(* IEC 61131-3 sources: NachHouse_TST/API/api_V12, 8 files *)

(* ---- _01_Types.ST ---- *)
// Konštanty určujú rozmery virtuálnej pamäte a počet typov ; Constants define virtual-memory dimensions and the number of data types.
VAR_GLOBAL CONSTANT
  _NH_ZONES {HIDDEN} : USINT := 5;      // Počet podporovaných pamäťových zón PLC ; Number of PLC memory zones used by this model.
  _NH_RAM {HIDDEN}   : UDINT := 10000;  // Veľkosť poľa mRam v bajtoch ; Size of the mRam byte array.
  _NH_CFG {HIDDEN}   : INT := 2;        // Počet typov registrovaných v aCfg ; Number of data types registered in aCfg.
END_VAR

// Nasledujú interné typy, dátové záznamy a dve publikované aplikačné štruktúry ; The following are internal types, data records, and two published application structures.
TYPE
  // Príznaky štartu a inicializácie programu ; Program startup and initialization flags.
  NH_SYS {HIDDEN}: STRUCT
    Ini     : INT := 250;    // Hodnota 250 povoľuje jednorazové naplnenie testovacích dát ; Value 250 enables the one-time test-data initialization.
    Restart : BOOL := TRUE;  // Označuje, že PLC práve štartuje ; Indicates that the PLC is starting.
  END_STRUCT;
  // Príklad spoločných identifikačných polí v oboch typoch ; Example of shared identification fields in both data types.
  NH_CFG_ALL {HIDDEN}: STRUCT
    RoomID     : INT := 12;  // Ukážkové ID miestnosti v spoločnej časti ; Sample room ID in the shared section.
    CategoryID : INT := 23;  // Ukážkové ID kategórie v spoločnej časti ; Sample category ID in the shared section.
  END_STRUCT;
  // Metaúdaje jedného typu: kód, veľkosť, počet viet a umiestnenie v mRam ; Metadata for one type: code, size, record count, and location in mRam.
  NH_CFG: STRUCT
    cfg     : STRING[4];                    // Kód typu, veľkosť vety, adresa, offset v mRam a počet viet ; Type code, record size, address, mRam offset, and record count.
    Siz     : UDINT;
    Ram     : UDINT;
    iRam    : UDINT;
    Rec     : UDINT;
    par     : USINT;                        // Pomocné klasifikačné a referenčné metadáta typu ; Auxiliary type classification and reference metadata.
    cat     : USINT;
    ref     : USINT := 251;
    ver     : USINT;
    tGrp    : USINT;                        // Klasifikačné údaje a veľkosti konfiguračnej/spoločnej časti ; Classification values and configuration/shared-section sizes.
    al      : USINT;
    cx      : UDINT;
    cf      : USINT := SIZEOF(NH_CFG_ALL);
    me      : UDINT;                        // Veľkosť stavovej časti, HW/I/O údaje a príznaky použiteľnosti ; State-section size, hardware/I/O data, and validity flags.
    hw      : USINT;
    io      : UDINT;
    Enabled : BOOL;
    ok      : BOOL;
  END_STRUCT;
  // Spoločné polia hlavičky každého záznamu ; Shared header fields for every record.
  NH_REC_ALL {HIDDEN}: STRUCT
    Ok : BOOL := TRUE;  // Príznak platnosti záznamu ; Record-validity flag.
    ID : INT;           // Identifikátor záznamu ; Record identifier.
  END_STRUCT;
  // Premenné živého stavu miestnosti uložené v časti mem ; Live room-state fields stored in the mem section.
  NH_ROOM_MEM: STRUCT
    rec          : NH_REC_ALL;  // Hlavička vety a spoločné identifikačné údaje ; Record header and shared identification data.
    all          : NH_CFG_ALL;
    Temperature  : REAL;        // Testovacie merania a stavové príznaky miestnosti ; Test measurements and room-state flags.
    Humidity     : REAL;
    Presence     : BOOL;
    DayPhase     : UINT;
    CategoryMask : DWORD;       // Maska kategórií, alarm a ďalšie binárne príznaky stavu ; Category mask, alarm level, and additional Boolean state flags.
    AlarmLevel   : USINT;
    Online       : BOOL;
    Twilight     : BOOL;
  END_STRUCT;
  // Konfiguračná časť miestnosti ; testovacie polia pokrývajú rôzne IEC typy ; Room configuration ; test fields cover different IEC data types.
  NH_ROOM_CFG: STRUCT
    Name           : STRING[32];                              // Názov a testovacie celé čísla so znamienkom aj bez neho ; Name and signed/unsigned integer test values.
    _Dint          : DINT;
    _Sint          : SINT;
    _Usint         : USINT;
    _Uint          : UINT;                                    // Testovacie 16-bitové a plávajúce čísla a krátky reťazec ; 16-bit and floating-point test values plus a short string.
    _Real          : REAL;
    _LReal         : LREAL;
    _String        : STRING[30];
    _StringCZSK    : STRING := 'SVKBEGIN_+ľščťžýáíé_SVKEND';  // Reťazec s diakritikou overuje prevod CP1250 na UTF-8 a späť ; A diacritic-bearing string tests conversion between CP1250 and UTF-8.
    _BYTE          : BYTE;                                    // Testovacie bajtové a časové typy ; Byte-sized and date/time test types.
    _WORD          : WORD;
    _TIME          : TIME;
    _DATE          : DATE;
    _TIME_OF_DAY   : TOD;                                     // Testovacie typy času dňa a dátumu s časom ; Test values for time-of-day and date-time types.
    _DATE_AND_TIME : DT;
  END_STRUCT;
  // Celá verejná veta miestnosti spája živý stav a konfiguráciu ; One public room record combines live state and configuration.
  NH_ROOM {PUBLIC}: STRUCT
    mem : NH_ROOM_MEM;  // Podštruktúra prevádzkového stavu miestnosti ; Nested room operating-state structure.
    cfg : NH_ROOM_CFG;  // Podštruktúra konfiguračných hodnôt miestnosti ; Nested room-configuration structure.
  END_STRUCT;
  // Živý stav používateľa oddelený od jeho konfigurácie ; Live user state separated from user configuration.
  NH_USERS_MEM: STRUCT
    rec        : NH_REC_ALL;  // Hlavička, spoločné identifikátory a stav pripojenia ; Header, shared identifiers, and connection state.
    all        : NH_CFG_ALL;
    Connected  : BOOL;
    LastError  : STRING[80];  // Posledná chyba a časová značka poslednej aktualizácie ; Last error and timestamp of the latest update.
    LastUpdate : UDINT;
  END_STRUCT;
  // Konfigurácia používateľa vrátane práv, zón, IP a ďalších polí ; User configuration including rights, zones, IP addresses, and other fields.
  NH_USERS_CFG: STRUCT
    Name       : STRING[32];                                                                                                              // Meno používateľa a predvoľby úvodnej obrazovky ; User name and home-screen preferences.
    LoginHome  : BOOL := TRUE;
    DshSet     : BOOL := FALSE;
    OwnDSH     : BOOL := TRUE;                                                                                                            // Príznaky vlastných obrazoviek a úroveň oprávnenia ; Custom-screen flags and access-right level.
    OwnQCK     : BOOL := TRUE;
    UsrRight   : USINT := 1;
    ZonList    : ARRAY[1..16] OF BOOL := [1, 1, 1, 1, 1, 1, 1, 1, 1, 1, 1, 1, 1, 1, 1, 1];                                                // Prístup používateľa k šestnástim zónam ; User access flags for sixteen zones.
    sbj        : USINT := 1;                                                                                                              // Predmet, jazyk a osem obľúbených položiek ; Subject, language, and eight favorites.
    lng        : USINT;
    fav        : ARRAY[0..7] OF USINT;
    keyPas     : STRING[6];                                                                                                               // Krátky testovací kľúč, počet IP adries a tri adresy ; Test key, IP-address count, and three addresses.
    IPnbr      : USINT := 1;
    IP         : ARRAY[1..3] OF STRING[15];
    mail       : STRING[50];                                                                                                              // Kontaktný e-mail a testovacie autorizačné tokeny ; Contact email and test authorization tokens.
    TOKENAPPLE : STRING[90];
    TOKENUNI   : STRING[100];
    gsm        : STRING[15];                                                                                                              // Telefón, vzhľad a osem príznakov správ ; Phone, appearance, and eight message flags.
    skin       : USINT;
    msg        : ARRAY[0..7] OF BOOL;
    Brw        : ARRAY[0..30] OF USINT := [0, 1, 1, 1, 1, 1, 1, 1, 1, 1, 1, 1, 1, 1, 1, 1, 1, 1, 1, 1, 1, 1, 1, 1, 1, 1, 1, 1, 1, 1, 1];  // Tridsaťjeden testovacích hodnôt pre prehliadač ; Thirty-one test values for browser-related settings.
  END_STRUCT;
  // Celá verejná veta používateľa spája stav a konfiguráciu ; One public user record combines state and configuration.
  NH_USER {PUBLIC}: STRUCT
    mem : NH_USERS_MEM;
    cfg : NH_USERS_CFG;
  END_STRUCT;
END_TYPE

VAR_GLOBAL
  mRam : ARRAY[0.._NH_RAM] OF BYTE;        // Spoločný bajtový priestor, v ktorom sú uložené všetky vety ; Shared byte-addressable memory containing all records.
  aSys : NH_SYS;                           // Stavové príznaky inicializácie programu ; Program initialization state.
  aCfg : ARRAY[1.._NH_CFG] OF NH_CFG := [  // Tabuľka typov: určuje ich veľkosti, počty viet a rozloženie v mRam ; Type table: defines sizes, record counts, and placement in mRam.
    (cfg := 'ROOM', Enabled := TRUE, ver := 1, Siz := SIZEOF(NH_ROOM),
     Rec := 10, cx := SIZEOF(NH_ROOM.cfg), me := SIZEOF(NH_ROOM.mem)),
    (cfg := 'USER', Enabled := TRUE, ver := 1, Siz := SIZEOF(NH_USER),
     Rec := 10, cx := SIZEOF(NH_USER.cfg), me := SIZEOF(NH_USER.mem),
     cat := 31, ref := 254)
  ];
  xRoom : PTR_TO NH_ROOM;  // Ukazovateľ na začiatok poľa viet ROOM v mRam ; Pointer to the first ROOM record in mRam.
  xUser : PTR_TO NH_USER;  // Ukazovateľ na začiatok poľa viet USER v mRam ; Pointer to the first USER record in mRam.

  yRooms : ARRAY[1..10] OF NH_ROOM;  // Iba zdroj testovacích dát ; po skopírovaní do mRam sa ďalej nepoužíva. ; Test-data source only ; unused after copying into mRam.
  yUsers : ARRAY[1..10] OF NH_USER;  // Zdroj testovacích viet USER ; po skopírovaní do mRam sa ďalej nepoužíva ; Source of USER test records ; unused after copying into mRam.

  DepRq {PUBLIC_API}   : BOOL := FALSE;        // Požiadavka na aktiváciu balíka ; Package-activation request.
  DepRes {PUBLIC_API}  : USINT := 0;           // Výsledkový kód aktivácie balíka ; Package-activation result code.
  BuildNo {PUBLIC_API} : UDINT := 2026100726;  // Číslo zostavenia na kontrolu nasadenej verzie ; Build number used to verify the deployed version.

  TxCf {PUBLIC_API}   : USINT := 2;  // Klient nastaví typ a vetu ; TxRq ako posledné spustí export. Nula znamená všetky vety. ; The client sets type and record ; TxRq starts the export last. Zero means all records.
  TxRec {PUBLIC_API}  : UDINT := 0;  // Číslo exportovanej vety ; nula znamená všetky vety vybraného typu ; Record to export ; zero means all records of the selected type.
  TxRq {PUBLIC_API}   : UDINT := 1;  // Klient zmenou čísla spustí nový export ; A new value starts an export request.
  TxDone {PUBLIC_API} : UDINT := 0;  // Potvrdí číslo dokončenej požiadavky na export ; Echoes the completed export request number.
  TxErr {PUBLIC_API}  : USINT := 0;  // Nula znamená úspech ; nenulová hodnota označuje chybu exportu ; Zero means success ; nonzero indicates an export error.

  RxRq    {PUBLIC_API} : UDINT := 0;  // Po prijatí rx.json klient zapíše nové RxRq a tým spustí jeho import. ; After rx.json is received, the client writes a new RxRq to start its import.
  RxDone  {PUBLIC_API} : UDINT := 0;  // Potvrdí číslo dokončenej požiadavky na import ; Echoes the completed import request number.
  RxErr   {PUBLIC_API} : USINT := 0;  // Nula znamená úspešný import ; inak obsahuje kód chyby ; Zero means import succeeded ; otherwise contains an error code.

  rxBuf   {PUBLIC_API} : ARRAY[0..63] OF DWORD;  // Jeden blok klienta má 64 DWORD, teda kapacitu 256 bajtov. ; One client block contains 64 DWORD values, providing 256 bytes of capacity. ; Klient zapíše dáta a metadáta ; RbRq mení až po nich. ; The client writes data and metadata first, then changes RbRq.
  RbOfs   {PUBLIC_API} : UDINT := 0;             // Offset bloku v celom súbore ; Block offset within the complete file.
  RbLen   {PUBLIC_API} : UINT := 0;              // Počet platných bajtov v tomto bloku ; Number of valid bytes in this block.
  RbTotal {PUBLIC_API} : UDINT := 0;             // Celková veľkosť prijímaného súboru ; Total size of the incoming file.
  RbCrc   {PUBLIC_API} : DWORD := 0;             // Očakávaný CRC32 súčet celého súboru ; Expected CRC32 checksum of the complete file.
  RbRq    {PUBLIC_API} : UDINT := 0;             // Spúšťací čítač bloku ; klient ho zapisuje až po dátach ; Block trigger counter ; written only after the block data.
  RbAck   {PUBLIC_API} : UDINT := 0;             // Potvrdzuje spracované číslo bloku ; Acknowledges the processed block number.
  RbWrote {PUBLIC_API} : UDINT := 0;             // Počet bajtov už uložených do rx.json ; Number of bytes already written to rx.json.
  RbReady {PUBLIC_API} : BOOL := FALSE;          // TRUE znamená celý súbor uložený a CRC overené ; TRUE means the full file is written and its CRC is valid.
  RbErr   {PUBLIC_API} : USINT := 0;             // Výsledok posledného bloku ; nula znamená úspech ; Result of the latest block ; zero means success.
END_VAR

(* ---- _03_Schema.ST ---- *)
// Automaticky vygenerované z api_V12.pux ; neupravovať ručne. ; GENERATED from api_V12.pux. Do not edit manually.
VAR_GLOBAL CONSTANT
  SCH_BOOL          : USINT := 16#01;        // Kód typu BOOL v schéme ; BOOL type code in the schema
  SCH_SINT          : USINT := 16#02;        // Kód typu SINT v schéme ; SINT type code in the schema
  SCH_USINT         : USINT := 16#03;        // Kód typu USINT v schéme ; USINT type code in the schema
  SCH_INT           : USINT := 16#04;        // Kód typu INT v schéme ; INT type code in the schema
  SCH_UINT          : USINT := 16#05;        // Kód typu UINT v schéme ; UINT type code in the schema
  SCH_DINT          : USINT := 16#06;        // Kód typu DINT v schéme ; DINT type code in the schema
  SCH_UDINT         : USINT := 16#07;        // Kód typu UDINT v schéme ; UDINT type code in the schema
  SCH_BYTE          : USINT := 16#08;        // Kód typu BYTE v schéme ; BYTE type code in the schema
  SCH_WORD          : USINT := 16#09;        // Kód typu WORD v schéme ; WORD type code in the schema
  SCH_DWORD         : USINT := 16#0A;        // Kód typu DWORD v schéme ; DWORD type code in the schema
  SCH_REAL          : USINT := 16#0B;        // Kód typu REAL v schéme ; REAL type code in the schema
  SCH_LREAL         : USINT := 16#0C;        // Kód typu LREAL v schéme ; LREAL type code in the schema
  SCH_STRING        : USINT := 16#0D;        // Kód reťazca v schéme ; String type code in the schema
  SCH_TIME          : USINT := 16#0E;        // Kód typu TIME v schéme ; TIME type code in the schema
  SCH_DATE          : USINT := 16#0F;        // Kód typu DATE v schéme ; DATE type code in the schema
  SCH_TIME_OF_DAY   : USINT := 16#10;        // Kód typu TOD v schéme ; TOD type code in the schema
  SCH_DATE_AND_TIME : USINT := 16#11;        // Kód typu DT v schéme ; DT type code in the schema
  SCH_STRUCT        : USINT := 16#12;        // Kód vnorenej štruktúry v schéme ; Nested-structure type code in the schema
  SCH_ARRAY         : USINT := 16#80;        // Príznak poľa kombinovaný so základným typom ; Array flag combined with the base type
  SCH_BASE          : USINT := 16#7F;        // Maska na získanie základného typu ; Mask used to extract the base type
  SCH_DEF_N         : UINT := 2;             // Počet definovaných aplikačných typov ; Number of application types defined
  SCH_NODE_N        : UINT := 62;            // Počet uzlov stromu štruktúr ; Number of structure-tree nodes
  SCH_LEAF_N        : UINT := 115;           // Počet úplných ciest k položkám ; Number of complete field paths
  SCH_PUX_CRC       : DWORD := 16#B72908B3;  // Kontrolný súčet zdrojového PUX ; Checksum of the source PUX
END_VAR

TYPE
  NH_SCH : STRUCT
    Cfg  : USINT;       // Poradové číslo typu v aCfg ; Type index in aCfg
    Code : STRING[4];   // Kód typu používaný v JSON obálke ; Type code used in the JSON envelope
    Nam  : STRING[16];  // Názov typu alebo uzla podľa kontextu ; Type or node name, depending on context
    Siz  : UDINT;       // Veľkosť jednej celej vety v bajtoch ; Size of one complete record in bytes
    Fst  : UINT;        // Index prvého uzla typu ; Index of the first node for this type
    Cnt  : UINT;        // Počet uzlov typu ; Number of nodes for this type
    LFst : UINT;        // Index prvej úplnej cesty poľa ; Index of the first complete field path
    LCnt : UINT;        // Počet úplných ciest poľa ; Number of complete field paths
  END_STRUCT;
  NH_NODE : STRUCT
    Nam  : STRING[14];  // Názov typu alebo uzla podľa kontextu ; Type or node name, depending on context
    Tag  : USINT;       // Kód dátového typu a prípadný príznak poľa ; Data-type code and optional array flag
    Ofs  : UINT;        // Offset položky od začiatku rodiča ; Field offset from the parent start
    Span : UINT;        // Veľkosť položky v bajtoch ; Field size in bytes
    Aux  : UINT;        // Doplnkový údaj podľa typu uzla ; Auxiliary value interpreted by node type
    Cnt  : UINT;        // Počet uzlov typu ; Number of nodes for this type
    Lo   : INT;         // Dolná hranica poľa ; Array lower bound
  END_STRUCT;
  NH_LEAF : STRUCT
    Pth    : STRING[18];  // Úplná cesta poľa od koreňa vety ; Complete field path from the record root
    Tag    : USINT;       // Kód dátového typu a prípadný príznak poľa ; Data-type code and optional array flag
    Ofs    : UINT;        // Offset položky od začiatku rodiča ; Field offset from the parent start
    Span   : UINT;        // Veľkosť položky v bajtoch ; Field size in bytes
    BitPos : SINT;        // Pozícia BOOL poľa v bajte ; BOOL field bit position within its byte
  END_STRUCT;
END_TYPE

VAR_GLOBAL
  aSch : ARRAY[1..2] OF NH_SCH := [  // Tabuľka rozsahov uzlov a polí pre každý typ ; Per-type ranges of nodes and fields
    (Cfg := 1, Code := 'ROOM', Nam := 'NH_ROOM', Siz := 216, Fst := 1, Cnt := 31, LFst := 1, LCnt := 27),
    (Cfg := 2, Code := 'USER', Nam := 'NH_USER', Siz := 488, Fst := 32, Cnt := 31, LFst := 28, LCnt := 88)
  ];
  aNode : ARRAY[1..62] OF NH_NODE := [  // Sploštený strom všetkých uzlov štruktúr ; Flattened tree of all structure nodes
    (Nam := 'mem', Tag := 16#12, Ofs := 0, Span := 24, Aux := 14, Cnt := 0, Lo := 0),
    (Nam := 'rec', Tag := 16#12, Ofs := 0, Span := 3, Aux := 2, Cnt := 0, Lo := 0),
    (Nam := 'Ok', Tag := 16#01, Ofs := 0, Span := 1, Aux := 0, Cnt := 0, Lo := 0),
    (Nam := 'ID', Tag := 16#04, Ofs := 1, Span := 2, Aux := 0, Cnt := 0, Lo := 0),
    (Nam := 'all', Tag := 16#12, Ofs := 3, Span := 4, Aux := 2, Cnt := 0, Lo := 0),
    (Nam := 'RoomID', Tag := 16#04, Ofs := 0, Span := 2, Aux := 0, Cnt := 0, Lo := 0),
    (Nam := 'CategoryID', Tag := 16#04, Ofs := 2, Span := 2, Aux := 0, Cnt := 0, Lo := 0),
    (Nam := 'Temperature', Tag := 16#0B, Ofs := 7, Span := 4, Aux := 0, Cnt := 0, Lo := 0),
    (Nam := 'Humidity', Tag := 16#0B, Ofs := 11, Span := 4, Aux := 0, Cnt := 0, Lo := 0),
    (Nam := 'Presence', Tag := 16#01, Ofs := 15, Span := 1, Aux := 0, Cnt := 0, Lo := 0),
    (Nam := 'DayPhase', Tag := 16#05, Ofs := 16, Span := 2, Aux := 0, Cnt := 0, Lo := 0),
    (Nam := 'CategoryMask', Tag := 16#0A, Ofs := 18, Span := 4, Aux := 0, Cnt := 0, Lo := 0),
    (Nam := 'AlarmLevel', Tag := 16#03, Ofs := 22, Span := 1, Aux := 0, Cnt := 0, Lo := 0),
    (Nam := 'Online', Tag := 16#01, Ofs := 23, Span := 1, Aux := 0, Cnt := 0, Lo := 0),
    (Nam := 'Twilight', Tag := 16#01, Ofs := 23, Span := 1, Aux := 1, Cnt := 0, Lo := 0),
    (Nam := 'cfg', Tag := 16#12, Ofs := 24, Span := 192, Aux := 15, Cnt := 0, Lo := 0),
    (Nam := 'Name', Tag := 16#0D, Ofs := 0, Span := 33, Aux := 0, Cnt := 0, Lo := 0),
    (Nam := '_Dint', Tag := 16#06, Ofs := 33, Span := 4, Aux := 0, Cnt := 0, Lo := 0),
    (Nam := '_Sint', Tag := 16#02, Ofs := 37, Span := 1, Aux := 0, Cnt := 0, Lo := 0),
    (Nam := '_Usint', Tag := 16#03, Ofs := 38, Span := 1, Aux := 0, Cnt := 0, Lo := 0),
    (Nam := '_Uint', Tag := 16#05, Ofs := 39, Span := 2, Aux := 0, Cnt := 0, Lo := 0),
    (Nam := '_Real', Tag := 16#0B, Ofs := 41, Span := 4, Aux := 0, Cnt := 0, Lo := 0),
    (Nam := '_LReal', Tag := 16#0C, Ofs := 45, Span := 8, Aux := 0, Cnt := 0, Lo := 0),
    (Nam := '_String', Tag := 16#0D, Ofs := 53, Span := 31, Aux := 0, Cnt := 0, Lo := 0),
    (Nam := '_StringCZSK', Tag := 16#0D, Ofs := 84, Span := 81, Aux := 0, Cnt := 0, Lo := 0),
    (Nam := '_BYTE', Tag := 16#08, Ofs := 165, Span := 1, Aux := 0, Cnt := 0, Lo := 0),
    (Nam := '_WORD', Tag := 16#09, Ofs := 166, Span := 2, Aux := 0, Cnt := 0, Lo := 0),
    (Nam := '_TIME', Tag := 16#0E, Ofs := 168, Span := 4, Aux := 0, Cnt := 0, Lo := 0),
    (Nam := '_DATE', Tag := 16#0F, Ofs := 172, Span := 8, Aux := 0, Cnt := 0, Lo := 0),
    (Nam := '_TIME_OF_DAY', Tag := 16#10, Ofs := 180, Span := 4, Aux := 0, Cnt := 0, Lo := 0),
    (Nam := '_DATE_AND_TIME', Tag := 16#11, Ofs := 184, Span := 8, Aux := 0, Cnt := 0, Lo := 0),
    (Nam := 'mem', Tag := 16#12, Ofs := 0, Span := 93, Aux := 9, Cnt := 0, Lo := 0),
    (Nam := 'rec', Tag := 16#12, Ofs := 0, Span := 3, Aux := 2, Cnt := 0, Lo := 0),
    (Nam := 'Ok', Tag := 16#01, Ofs := 0, Span := 1, Aux := 0, Cnt := 0, Lo := 0),
    (Nam := 'ID', Tag := 16#04, Ofs := 1, Span := 2, Aux := 0, Cnt := 0, Lo := 0),
    (Nam := 'all', Tag := 16#12, Ofs := 3, Span := 4, Aux := 2, Cnt := 0, Lo := 0),
    (Nam := 'RoomID', Tag := 16#04, Ofs := 0, Span := 2, Aux := 0, Cnt := 0, Lo := 0),
    (Nam := 'CategoryID', Tag := 16#04, Ofs := 2, Span := 2, Aux := 0, Cnt := 0, Lo := 0),
    (Nam := 'Connected', Tag := 16#01, Ofs := 7, Span := 1, Aux := 0, Cnt := 0, Lo := 0),
    (Nam := 'LastError', Tag := 16#0D, Ofs := 8, Span := 81, Aux := 0, Cnt := 0, Lo := 0),
    (Nam := 'LastUpdate', Tag := 16#07, Ofs := 89, Span := 4, Aux := 0, Cnt := 0, Lo := 0),
    (Nam := 'cfg', Tag := 16#12, Ofs := 93, Span := 395, Aux := 20, Cnt := 0, Lo := 0),
    (Nam := 'Name', Tag := 16#0D, Ofs := 0, Span := 33, Aux := 0, Cnt := 0, Lo := 0),
    (Nam := 'LoginHome', Tag := 16#01, Ofs := 33, Span := 1, Aux := 0, Cnt := 0, Lo := 0),
    (Nam := 'DshSet', Tag := 16#01, Ofs := 33, Span := 1, Aux := 1, Cnt := 0, Lo := 0),
    (Nam := 'OwnDSH', Tag := 16#01, Ofs := 33, Span := 1, Aux := 2, Cnt := 0, Lo := 0),
    (Nam := 'OwnQCK', Tag := 16#01, Ofs := 33, Span := 1, Aux := 3, Cnt := 0, Lo := 0),
    (Nam := 'UsrRight', Tag := 16#03, Ofs := 34, Span := 1, Aux := 0, Cnt := 0, Lo := 0),
    (Nam := 'ZonList', Tag := 16#81, Ofs := 35, Span := 2, Aux := 0, Cnt := 16, Lo := 1),
    (Nam := 'sbj', Tag := 16#03, Ofs := 37, Span := 1, Aux := 0, Cnt := 0, Lo := 0),
    (Nam := 'lng', Tag := 16#03, Ofs := 38, Span := 1, Aux := 0, Cnt := 0, Lo := 0),
    (Nam := 'fav', Tag := 16#83, Ofs := 39, Span := 8, Aux := 1, Cnt := 8, Lo := 0),
    (Nam := 'keyPas', Tag := 16#0D, Ofs := 47, Span := 7, Aux := 0, Cnt := 0, Lo := 0),
    (Nam := 'IPnbr', Tag := 16#03, Ofs := 54, Span := 1, Aux := 0, Cnt := 0, Lo := 0),
    (Nam := 'IP', Tag := 16#8D, Ofs := 55, Span := 48, Aux := 16, Cnt := 3, Lo := 1),
    (Nam := 'mail', Tag := 16#0D, Ofs := 103, Span := 51, Aux := 0, Cnt := 0, Lo := 0),
    (Nam := 'TOKENAPPLE', Tag := 16#0D, Ofs := 154, Span := 91, Aux := 0, Cnt := 0, Lo := 0),
    (Nam := 'TOKENUNI', Tag := 16#0D, Ofs := 245, Span := 101, Aux := 0, Cnt := 0, Lo := 0),
    (Nam := 'gsm', Tag := 16#0D, Ofs := 346, Span := 16, Aux := 0, Cnt := 0, Lo := 0),
    (Nam := 'skin', Tag := 16#03, Ofs := 362, Span := 1, Aux := 0, Cnt := 0, Lo := 0),
    (Nam := 'msg', Tag := 16#81, Ofs := 363, Span := 1, Aux := 0, Cnt := 8, Lo := 0),
    (Nam := 'Brw', Tag := 16#83, Ofs := 364, Span := 31, Aux := 1, Cnt := 31, Lo := 0)
  ];
  aLeaf : ARRAY[1..115] OF NH_LEAF := [  // Tabuľka úplných názvov koncových polí ; Lookup table of complete leaf-field names
    (Pth := 'mem.rec.Ok', Tag := 16#01, Ofs := 0, Span := 1, BitPos := 0),
    (Pth := 'mem.rec.ID', Tag := 16#04, Ofs := 1, Span := 2, BitPos := -1),
    (Pth := 'mem.all.RoomID', Tag := 16#04, Ofs := 3, Span := 2, BitPos := -1),
    (Pth := 'mem.all.CategoryID', Tag := 16#04, Ofs := 5, Span := 2, BitPos := -1),
    (Pth := 'mem.Temperature', Tag := 16#0B, Ofs := 7, Span := 4, BitPos := -1),
    (Pth := 'mem.Humidity', Tag := 16#0B, Ofs := 11, Span := 4, BitPos := -1),
    (Pth := 'mem.Presence', Tag := 16#01, Ofs := 15, Span := 1, BitPos := 0),
    (Pth := 'mem.DayPhase', Tag := 16#05, Ofs := 16, Span := 2, BitPos := -1),
    (Pth := 'mem.CategoryMask', Tag := 16#0A, Ofs := 18, Span := 4, BitPos := -1),
    (Pth := 'mem.AlarmLevel', Tag := 16#03, Ofs := 22, Span := 1, BitPos := -1),
    (Pth := 'mem.Online', Tag := 16#01, Ofs := 23, Span := 1, BitPos := 0),
    (Pth := 'mem.Twilight', Tag := 16#01, Ofs := 23, Span := 1, BitPos := 1),
    (Pth := 'cfg.Name', Tag := 16#0D, Ofs := 24, Span := 33, BitPos := -1),
    (Pth := 'cfg._Dint', Tag := 16#06, Ofs := 57, Span := 4, BitPos := -1),
    (Pth := 'cfg._Sint', Tag := 16#02, Ofs := 61, Span := 1, BitPos := -1),
    (Pth := 'cfg._Usint', Tag := 16#03, Ofs := 62, Span := 1, BitPos := -1),
    (Pth := 'cfg._Uint', Tag := 16#05, Ofs := 63, Span := 2, BitPos := -1),
    (Pth := 'cfg._Real', Tag := 16#0B, Ofs := 65, Span := 4, BitPos := -1),
    (Pth := 'cfg._LReal', Tag := 16#0C, Ofs := 69, Span := 8, BitPos := -1),
    (Pth := 'cfg._String', Tag := 16#0D, Ofs := 77, Span := 31, BitPos := -1),
    (Pth := 'cfg._StringCZSK', Tag := 16#0D, Ofs := 108, Span := 81, BitPos := -1),
    (Pth := 'cfg._BYTE', Tag := 16#08, Ofs := 189, Span := 1, BitPos := -1),
    (Pth := 'cfg._WORD', Tag := 16#09, Ofs := 190, Span := 2, BitPos := -1),
    (Pth := 'cfg._TIME', Tag := 16#0E, Ofs := 192, Span := 4, BitPos := -1),
    (Pth := 'cfg._DATE', Tag := 16#0F, Ofs := 196, Span := 8, BitPos := -1),
    (Pth := 'cfg._TIME_OF_DAY', Tag := 16#10, Ofs := 204, Span := 4, BitPos := -1),
    (Pth := 'cfg._DATE_AND_TIME', Tag := 16#11, Ofs := 208, Span := 8, BitPos := -1),
    (Pth := 'mem.rec.Ok', Tag := 16#01, Ofs := 0, Span := 1, BitPos := 0),
    (Pth := 'mem.rec.ID', Tag := 16#04, Ofs := 1, Span := 2, BitPos := -1),
    (Pth := 'mem.all.RoomID', Tag := 16#04, Ofs := 3, Span := 2, BitPos := -1),
    (Pth := 'mem.all.CategoryID', Tag := 16#04, Ofs := 5, Span := 2, BitPos := -1),
    (Pth := 'mem.Connected', Tag := 16#01, Ofs := 7, Span := 1, BitPos := 0),
    (Pth := 'mem.LastError', Tag := 16#0D, Ofs := 8, Span := 81, BitPos := -1),
    (Pth := 'mem.LastUpdate', Tag := 16#07, Ofs := 89, Span := 4, BitPos := -1),
    (Pth := 'cfg.Name', Tag := 16#0D, Ofs := 93, Span := 33, BitPos := -1),
    (Pth := 'cfg.LoginHome', Tag := 16#01, Ofs := 126, Span := 1, BitPos := 0),
    (Pth := 'cfg.DshSet', Tag := 16#01, Ofs := 126, Span := 1, BitPos := 1),
    (Pth := 'cfg.OwnDSH', Tag := 16#01, Ofs := 126, Span := 1, BitPos := 2),
    (Pth := 'cfg.OwnQCK', Tag := 16#01, Ofs := 126, Span := 1, BitPos := 3),
    (Pth := 'cfg.UsrRight', Tag := 16#03, Ofs := 127, Span := 1, BitPos := -1),
    (Pth := 'cfg.ZonList[0]', Tag := 16#01, Ofs := 128, Span := 1, BitPos := 0),
    (Pth := 'cfg.ZonList[1]', Tag := 16#01, Ofs := 128, Span := 1, BitPos := 1),
    (Pth := 'cfg.ZonList[2]', Tag := 16#01, Ofs := 128, Span := 1, BitPos := 2),
    (Pth := 'cfg.ZonList[3]', Tag := 16#01, Ofs := 128, Span := 1, BitPos := 3),
    (Pth := 'cfg.ZonList[4]', Tag := 16#01, Ofs := 128, Span := 1, BitPos := 4),
    (Pth := 'cfg.ZonList[5]', Tag := 16#01, Ofs := 128, Span := 1, BitPos := 5),
    (Pth := 'cfg.ZonList[6]', Tag := 16#01, Ofs := 128, Span := 1, BitPos := 6),
    (Pth := 'cfg.ZonList[7]', Tag := 16#01, Ofs := 128, Span := 1, BitPos := 7),
    (Pth := 'cfg.ZonList[8]', Tag := 16#01, Ofs := 129, Span := 1, BitPos := 0),
    (Pth := 'cfg.ZonList[9]', Tag := 16#01, Ofs := 129, Span := 1, BitPos := 1),
    (Pth := 'cfg.ZonList[10]', Tag := 16#01, Ofs := 129, Span := 1, BitPos := 2),
    (Pth := 'cfg.ZonList[11]', Tag := 16#01, Ofs := 129, Span := 1, BitPos := 3),
    (Pth := 'cfg.ZonList[12]', Tag := 16#01, Ofs := 129, Span := 1, BitPos := 4),
    (Pth := 'cfg.ZonList[13]', Tag := 16#01, Ofs := 129, Span := 1, BitPos := 5),
    (Pth := 'cfg.ZonList[14]', Tag := 16#01, Ofs := 129, Span := 1, BitPos := 6),
    (Pth := 'cfg.ZonList[15]', Tag := 16#01, Ofs := 129, Span := 1, BitPos := 7),
    (Pth := 'cfg.sbj', Tag := 16#03, Ofs := 130, Span := 1, BitPos := -1),
    (Pth := 'cfg.lng', Tag := 16#03, Ofs := 131, Span := 1, BitPos := -1),
    (Pth := 'cfg.fav[0]', Tag := 16#03, Ofs := 132, Span := 1, BitPos := -1),
    (Pth := 'cfg.fav[1]', Tag := 16#03, Ofs := 133, Span := 1, BitPos := -1),
    (Pth := 'cfg.fav[2]', Tag := 16#03, Ofs := 134, Span := 1, BitPos := -1),
    (Pth := 'cfg.fav[3]', Tag := 16#03, Ofs := 135, Span := 1, BitPos := -1),
    (Pth := 'cfg.fav[4]', Tag := 16#03, Ofs := 136, Span := 1, BitPos := -1),
    (Pth := 'cfg.fav[5]', Tag := 16#03, Ofs := 137, Span := 1, BitPos := -1),
    (Pth := 'cfg.fav[6]', Tag := 16#03, Ofs := 138, Span := 1, BitPos := -1),
    (Pth := 'cfg.fav[7]', Tag := 16#03, Ofs := 139, Span := 1, BitPos := -1),
    (Pth := 'cfg.keyPas', Tag := 16#0D, Ofs := 140, Span := 7, BitPos := -1),
    (Pth := 'cfg.IPnbr', Tag := 16#03, Ofs := 147, Span := 1, BitPos := -1),
    (Pth := 'cfg.IP[0]', Tag := 16#0D, Ofs := 148, Span := 16, BitPos := -1),
    (Pth := 'cfg.IP[1]', Tag := 16#0D, Ofs := 164, Span := 16, BitPos := -1),
    (Pth := 'cfg.IP[2]', Tag := 16#0D, Ofs := 180, Span := 16, BitPos := -1),
    (Pth := 'cfg.mail', Tag := 16#0D, Ofs := 196, Span := 51, BitPos := -1),
    (Pth := 'cfg.TOKENAPPLE', Tag := 16#0D, Ofs := 247, Span := 91, BitPos := -1),
    (Pth := 'cfg.TOKENUNI', Tag := 16#0D, Ofs := 338, Span := 101, BitPos := -1),
    (Pth := 'cfg.gsm', Tag := 16#0D, Ofs := 439, Span := 16, BitPos := -1),
    (Pth := 'cfg.skin', Tag := 16#03, Ofs := 455, Span := 1, BitPos := -1),
    (Pth := 'cfg.msg[0]', Tag := 16#01, Ofs := 456, Span := 1, BitPos := 0),
    (Pth := 'cfg.msg[1]', Tag := 16#01, Ofs := 456, Span := 1, BitPos := 1),
    (Pth := 'cfg.msg[2]', Tag := 16#01, Ofs := 456, Span := 1, BitPos := 2),
    (Pth := 'cfg.msg[3]', Tag := 16#01, Ofs := 456, Span := 1, BitPos := 3),
    (Pth := 'cfg.msg[4]', Tag := 16#01, Ofs := 456, Span := 1, BitPos := 4),
    (Pth := 'cfg.msg[5]', Tag := 16#01, Ofs := 456, Span := 1, BitPos := 5),
    (Pth := 'cfg.msg[6]', Tag := 16#01, Ofs := 456, Span := 1, BitPos := 6),
    (Pth := 'cfg.msg[7]', Tag := 16#01, Ofs := 456, Span := 1, BitPos := 7),
    (Pth := 'cfg.Brw[0]', Tag := 16#03, Ofs := 457, Span := 1, BitPos := -1),
    (Pth := 'cfg.Brw[1]', Tag := 16#03, Ofs := 458, Span := 1, BitPos := -1),
    (Pth := 'cfg.Brw[2]', Tag := 16#03, Ofs := 459, Span := 1, BitPos := -1),
    (Pth := 'cfg.Brw[3]', Tag := 16#03, Ofs := 460, Span := 1, BitPos := -1),
    (Pth := 'cfg.Brw[4]', Tag := 16#03, Ofs := 461, Span := 1, BitPos := -1),
    (Pth := 'cfg.Brw[5]', Tag := 16#03, Ofs := 462, Span := 1, BitPos := -1),
    (Pth := 'cfg.Brw[6]', Tag := 16#03, Ofs := 463, Span := 1, BitPos := -1),
    (Pth := 'cfg.Brw[7]', Tag := 16#03, Ofs := 464, Span := 1, BitPos := -1),
    (Pth := 'cfg.Brw[8]', Tag := 16#03, Ofs := 465, Span := 1, BitPos := -1),
    (Pth := 'cfg.Brw[9]', Tag := 16#03, Ofs := 466, Span := 1, BitPos := -1),
    (Pth := 'cfg.Brw[10]', Tag := 16#03, Ofs := 467, Span := 1, BitPos := -1),
    (Pth := 'cfg.Brw[11]', Tag := 16#03, Ofs := 468, Span := 1, BitPos := -1),
    (Pth := 'cfg.Brw[12]', Tag := 16#03, Ofs := 469, Span := 1, BitPos := -1),
    (Pth := 'cfg.Brw[13]', Tag := 16#03, Ofs := 470, Span := 1, BitPos := -1),
    (Pth := 'cfg.Brw[14]', Tag := 16#03, Ofs := 471, Span := 1, BitPos := -1),
    (Pth := 'cfg.Brw[15]', Tag := 16#03, Ofs := 472, Span := 1, BitPos := -1),
    (Pth := 'cfg.Brw[16]', Tag := 16#03, Ofs := 473, Span := 1, BitPos := -1),
    (Pth := 'cfg.Brw[17]', Tag := 16#03, Ofs := 474, Span := 1, BitPos := -1),
    (Pth := 'cfg.Brw[18]', Tag := 16#03, Ofs := 475, Span := 1, BitPos := -1),
    (Pth := 'cfg.Brw[19]', Tag := 16#03, Ofs := 476, Span := 1, BitPos := -1),
    (Pth := 'cfg.Brw[20]', Tag := 16#03, Ofs := 477, Span := 1, BitPos := -1),
    (Pth := 'cfg.Brw[21]', Tag := 16#03, Ofs := 478, Span := 1, BitPos := -1),
    (Pth := 'cfg.Brw[22]', Tag := 16#03, Ofs := 479, Span := 1, BitPos := -1),
    (Pth := 'cfg.Brw[23]', Tag := 16#03, Ofs := 480, Span := 1, BitPos := -1),
    (Pth := 'cfg.Brw[24]', Tag := 16#03, Ofs := 481, Span := 1, BitPos := -1),
    (Pth := 'cfg.Brw[25]', Tag := 16#03, Ofs := 482, Span := 1, BitPos := -1),
    (Pth := 'cfg.Brw[26]', Tag := 16#03, Ofs := 483, Span := 1, BitPos := -1),
    (Pth := 'cfg.Brw[27]', Tag := 16#03, Ofs := 484, Span := 1, BitPos := -1),
    (Pth := 'cfg.Brw[28]', Tag := 16#03, Ofs := 485, Span := 1, BitPos := -1),
    (Pth := 'cfg.Brw[29]', Tag := 16#03, Ofs := 486, Span := 1, BitPos := -1),
    (Pth := 'cfg.Brw[30]', Tag := 16#03, Ofs := 487, Span := 1, BitPos := -1)
  ];
END_VAR

(* ---- _04_SchemaRun.ST ---- *)
// Stav validácie generovanej schémy ; Validation state for the generated schema.
VAR_GLOBAL
  SchOk    : BOOL := FALSE;  // TRUE až po úspešnej kontrole celej tabuľky schémy ; TRUE only after the entire schema table passes validation.
  SchErr   : USINT := 0;     // Kód prvej chyby zistený pri kontrole schémy ; First error code detected during schema validation.
  SchState : USINT := 0;     // Kontrola schémy sa vykoná raz a jej výsledok sa zapamätá ; Schema validation runs once and its result is cached. 0=new, 1=valid, 2=error
END_VAR

// Porovná vygenerovanú schému s aCfg a aktuálnym rozložením mRam. ; Compare the generated schema with aCfg and the current mRam layout.
// Overí počty, veľkosti, uzly a rozsahy schémy ešte pred prevodom ; Validate schema counts, sizes, nodes, and bounds before conversion.
FUNCTION SchInit : BOOL
  VAR
    Cf       : INT;                   // Index dátového typu v aCfg/aSch ; Data-type index in aCfg/aSch.
    Nd       : UINT;                  // Index práve kontrolovaného uzla štruktúry ; Index of the structure node being checked.
    Last     : UINT;                  // Posledný uzol patriaci aktuálnemu typu ; Last node belonging to the current type.
    Expected : UINT := 1;             // Očakávaný začiatok ďalšieho súvislého rozsahu uzlov ; Expected start of the next contiguous node range.
    BaseTag  : USINT;                 // Základný typ uzla po odobratí príznaku ARRAY ; Node base type after removing the ARRAY flag. ; Základný typ určuje výpočet prvku poľa ; The base type determines array-element addressing.
    NodeEnd  : UINT;                  // Koniec podstromu vnoreného STRUCT ; End of a nested STRUCT subtree.
    ElemSpan : UINT;                  // Veľkosť jedného prvku poľa STRUCT ; Size of one STRUCT-array element.
    Depth    : USINT;                 // Aktuálna hĺbka vnorenia pri kontrole uzlov ; Current nesting depth while validating nodes.
    EndStk   : ARRAY[0..15] OF UINT;  // Zásobník hraníc uzlov vnorených štruktúr ; Stack of node-range ends for nested structures.
    SpanStk  : ARRAY[0..15] OF UINT;  // Zásobník veľkostí rodičovských pamäťových oblastí ; Stack of parent memory-span sizes.
    RamEnd   : UDINT;                 // Koniec vyhradenej oblasti typu v mRam ; End of this type's reserved region in mRam.
  END_VAR

  SchInit := FALSE;
  // Použije zapamätaný úspech bez opakovania úplnej kontroly ; Reuse the cached success without repeating full validation.
  IF SchState = 1 THEN SchInit := TRUE; RETURN; END_IF;
  // Po predchádzajúcej chybe sa prevod bezpečne zastaví ; Stop conversion after a previously detected schema error.
  IF SchState = 2 THEN RETURN; END_IF;

  SchOk := FALSE;
  SchErr := 1;
  SchState := 2;
  IF SCH_DEF_N <> INT_TO_UINT(_NH_CFG) THEN RETURN; END_IF;

  // Porovná každý typ schémy s jeho konfiguráciou a rozložením v pamäti ; Compare each schema type with its configuration and memory layout.
  FOR Cf := 1 TO _NH_CFG DO
    IF aSch[Cf].Cfg <> INT_TO_USINT(Cf) THEN SchErr := 2; RETURN; END_IF;
    IF aSch[Cf].Code <> aCfg[Cf].cfg THEN SchErr := 3; RETURN; END_IF;
    IF aSch[Cf].Siz <> aCfg[Cf].Siz THEN SchErr := 4; RETURN; END_IF;
    IF (aSch[Cf].Fst <> Expected) OR (aSch[Cf].Cnt = 0) THEN SchErr := 5; RETURN; END_IF;
    Last := aSch[Cf].Fst + aSch[Cf].Cnt - 1;
    IF Last > SCH_NODE_N THEN SchErr := 6; RETURN; END_IF;
    Expected := Last + 1;

    RamEnd := aCfg[Cf].iRam + aCfg[Cf].Siz * aCfg[Cf].Rec;
    IF RamEnd > SIZEOF(mRam) THEN SchErr := 7; RETURN; END_IF;
    IF aCfg[Cf].Ram <> PTR_TO_UDINT(ADR(mRam[aCfg[Cf].iRam])) THEN SchErr := 8; RETURN; END_IF;

    Depth := 0;  // Začne kontrolu stromu uzlov od koreňa aktuálneho typu ; Start validating the node tree at the current type's root.
    EndStk[0] := Last + 1;
    SpanStk[0] := UDINT_TO_UINT(aSch[Cf].Siz);
    FOR Nd := aSch[Cf].Fst TO Last DO
      WHILE (Depth > 0) AND (Nd >= EndStk[Depth]) DO Depth := Depth - 1; END_WHILE;
      IF UINT_TO_UDINT(aNode[Nd].Ofs) + UINT_TO_UDINT(aNode[Nd].Span) > UINT_TO_UDINT(SpanStk[Depth]) THEN
        SchErr := 9; RETURN;
      END_IF;

      BaseTag := aNode[Nd].Tag MOD SCH_ARRAY;  // Oddelí základný dátový typ od príznaku poľa ; Separate the base data type from the array flag.
      IF (BaseTag < SCH_BOOL) OR (BaseTag > SCH_STRUCT) OR (aNode[Nd].Span = 0) THEN
        SchErr := 10; RETURN;
      END_IF;

      IF aNode[Nd].Tag >= SCH_ARRAY THEN
        IF aNode[Nd].Cnt = 0 THEN SchErr := 11; RETURN; END_IF;
        IF BaseTag = SCH_STRUCT THEN
          IF (aNode[Nd].Span MOD aNode[Nd].Cnt) <> 0 THEN SchErr := 12; RETURN; END_IF;
        ELSIF BaseTag = SCH_BOOL THEN
          IF (aNode[Nd].Aux + aNode[Nd].Cnt + 7) / 8 > aNode[Nd].Span THEN SchErr := 13; RETURN; END_IF;
        ELSE
          IF (aNode[Nd].Aux = 0) OR (aNode[Nd].Aux * aNode[Nd].Cnt <> aNode[Nd].Span) THEN
            SchErr := 14; RETURN;
          END_IF;
        END_IF;
      ELSE
        IF aNode[Nd].Cnt <> 0 THEN SchErr := 15; RETURN; END_IF;
        IF (BaseTag = SCH_BOOL) AND (aNode[Nd].Aux > 7) THEN SchErr := 16; RETURN; END_IF;
      END_IF;

      IF BaseTag = SCH_STRUCT THEN
        NodeEnd := Nd + 1 + aNode[Nd].Aux;
        IF NodeEnd > EndStk[Depth] THEN SchErr := 17; RETURN; END_IF;
        IF aNode[Nd].Aux > 0 THEN
          IF Depth >= 15 THEN SchErr := 18; RETURN; END_IF;
          IF aNode[Nd].Tag >= SCH_ARRAY THEN ElemSpan := aNode[Nd].Span / aNode[Nd].Cnt;
          ELSE ElemSpan := aNode[Nd].Span;
          END_IF;
          Depth := Depth + 1;
          EndStk[Depth] := NodeEnd;
          SpanStk[Depth] := ElemSpan;
        END_IF;
      END_IF;
    END_FOR;
  END_FOR;

  IF Expected <> SCH_NODE_N + 1 THEN SchErr := 19; RETURN; END_IF;
  SchErr := 0;  // Všetky kontroly prešli ; SchInit môže povoliť prevod ; All checks passed ; SchInit may allow conversion.
  SchOk := TRUE;
  SchState := 1;
  SchInit := TRUE;
END_FUNCTION

// Vráti začiatok zvolenej vety v mRam ; Rec sa čísluje od 1. ; Return the selected record's base address in mRam ; Rec is one-based.
// Vráti adresu vybranej vety v mRam alebo nulu pri neplatnom výbere ; Return the selected record's mRam address, or zero for an invalid selection.
FUNCTION SchRoot : UDINT
  VAR_INPUT
    Cf  : USINT;
    Rec : UDINT;
  END_VAR
  SchRoot := 0;
  IF NOT SchInit() THEN RETURN; END_IF;
  IF (Cf < 1) OR (Cf > UINT_TO_USINT(SCH_DEF_N)) THEN RETURN; END_IF;
  IF (Rec < 1) OR (Rec > aCfg[Cf].Rec) THEN RETURN; END_IF;
  IF NOT aCfg[Cf].Enabled OR NOT aCfg[Cf].ok THEN RETURN; END_IF;
  SchRoot := aCfg[Cf].Ram + (Rec - 1) * aCfg[Cf].Siz;
END_FUNCTION

// Vypočíta adresu uzla v rodičovi ; El pri poli je skutočný IEC index. ; Calculate a node address within its parent ; El is the actual IEC array index.
// Vypočíta adresu položky alebo prvku poľa z rodičovskej adresy a offsetu ; Calculate a field/array-element address from its parent and offset.
FUNCTION SchAdr : UDINT
  VAR_INPUT
    Parent : UDINT;
    Nd     : UINT;   // Index práve kontrolovaného uzla štruktúry ; Index of the structure node being checked.
    El     : INT;
  END_VAR
  VAR
    BaseTag : USINT;  // Základný typ uzla po odobratí príznaku ARRAY ; Node base type after removing the ARRAY flag. ; Základný typ určuje výpočet prvku poľa ; The base type determines array-element addressing.
    K       : UINT;   // Poradové číslo prvku od dolnej hranice poľa ; Zero-based element index from the array lower bound.
    BitPos  : UINT;   // Bitová pozícia BOOL prvku v bajte ; Bit position of a BOOL element within its byte.
  END_VAR
  SchAdr := 0;
  IF NOT SchInit() OR (Parent = 0) OR (Nd < 1) OR (Nd > SCH_NODE_N) THEN RETURN; END_IF;
  IF aNode[Nd].Tag < SCH_ARRAY THEN
    SchAdr := Parent + UINT_TO_UDINT(aNode[Nd].Ofs);
    RETURN;
  END_IF;
  IF (El < aNode[Nd].Lo) OR (El >= aNode[Nd].Lo + UINT_TO_INT(aNode[Nd].Cnt)) THEN RETURN; END_IF;
  K := INT_TO_UINT(El - aNode[Nd].Lo);
  BaseTag := aNode[Nd].Tag MOD SCH_ARRAY;
  IF BaseTag = SCH_BOOL THEN
    BitPos := aNode[Nd].Aux + K;
    SchAdr := Parent + UINT_TO_UDINT(aNode[Nd].Ofs) + UINT_TO_UDINT(BitPos / 8);
  ELSIF BaseTag = SCH_STRUCT THEN
    SchAdr := Parent + UINT_TO_UDINT(aNode[Nd].Ofs) + UINT_TO_UDINT(K * (aNode[Nd].Span / aNode[Nd].Cnt));
  ELSE
    SchAdr := Parent + UINT_TO_UDINT(aNode[Nd].Ofs) + UINT_TO_UDINT(K * aNode[Nd].Aux);
  END_IF;
END_FUNCTION

// Vráti bitovú pozíciu BOOL ; pri ostatných typoch vráti -1. ; Return the BOOL bit position, or -1 for other types.
// Vráti bitovú pozíciu BOOL ; pri inom type vráti -1 ; Return a BOOL bit position, or -1 for another type.
FUNCTION SchBit : SINT
  VAR_INPUT
    Nd : UINT;  // Index práve kontrolovaného uzla štruktúry ; Index of the structure node being checked.
    El : INT;
  END_VAR
  VAR
    K : UINT;  // Poradové číslo prvku od dolnej hranice poľa ; Zero-based element index from the array lower bound.
  END_VAR
  SchBit := -1;
  IF (Nd < 1) OR (Nd > SCH_NODE_N) THEN RETURN; END_IF;
  IF (aNode[Nd].Tag MOD SCH_ARRAY) <> SCH_BOOL THEN RETURN; END_IF;
  IF aNode[Nd].Tag < SCH_ARRAY THEN
    SchBit := UINT_TO_SINT(aNode[Nd].Aux);
    RETURN;
  END_IF;
  IF (El < aNode[Nd].Lo) OR (El >= aNode[Nd].Lo + UINT_TO_INT(aNode[Nd].Cnt)) THEN RETURN; END_IF;
  K := INT_TO_UINT(El - aNode[Nd].Lo);
  SchBit := UINT_TO_SINT((aNode[Nd].Aux + K) MOD 8);
END_FUNCTION

// Nájde ďalší uzol rovnakej úrovne a preskočí vnorený STRUCT. ; Find the next node at the same level, skipping a nested STRUCT.
// Vráti nasledujúci súrodenecký uzol a preskočí vnorený podstrom ; Return the next sibling node, skipping any nested subtree.
FUNCTION SchNext : UINT
  VAR_INPUT
    Nd : UINT;
  END_VAR
  SchNext := 0;
  IF (Nd < 1) OR (Nd > SCH_NODE_N) THEN RETURN; END_IF;
  IF (aNode[Nd].Tag MOD SCH_ARRAY) = SCH_STRUCT THEN SchNext := Nd + 1 + aNode[Nd].Aux;
  ELSE SchNext := Nd + 1;
  END_IF;
END_FUNCTION

(* ---- _05_TxJson.ST ---- *)
VAR_GLOBAL
  TxPath    : STRING[80] := '//RAM/tx.json';     // Cieľový súbor exportovaného JSON ; Destination file for exported JSON
  TxLogPath : STRING[80] := '//RAM/tx.log';      // Súbor meraní exportu ; Export measurement log file
  TxCRLF    : STRING[2] := '$0D$0A';             // Koniec riadka používaný v súbore ; Line ending used in the file
  TxH       : HANDLE := INVALID_HANDLE_VALUE;    // Handle otvoreného exportného súboru ; Handle of the open export file
  TxSeen    : UDINT := 0;                        // Posledná požiadavka už spracovaná PLC ; Latest request already processed by the PLC
  TxWorkErr : USINT := 0;                        // Pracovný kód chyby exportu ; Working export error code
  TxBytes   : UDINT := 0;                        // Počet bajtov zapísaných do súboru ; Number of bytes written to the file
  TxHex     : STRING[16] := '0123456789ABCDEF';  // Tabuľka číslic na zápis hexadecimálnych hodnôt ; Digit table for hexadecimal output
  TxSt      : USINT := 0;                        // Stavový automat exportu ; Export state-machine state
  TxCfW     : USINT := 0;                        // Typ vybraný pre aktuálny export ; Type selected for the current export
  TxFrom    : UDINT := 0;                        // Prvé číslo exportovanej vety ; First record number to export
  TxTo      : UDINT := 0;                        // Posledné číslo exportovanej vety ; Last record number to export
  TxNow     : UDINT := 0;                        // Číslo vety spracúvanej teraz ; Record number currently being processed
  TxRqW     : UDINT := 0;                        // Číslo požiadavky aktuálneho exportu ; Request number for the current export
  TxMode    : USINT := 0;                        // Režim výberu viet ; Record-selection mode ; 1=one, 2=range, 3=all
  TxMs0     : UDINT := 0;                        // Čas začiatku exportu v milisekundách ; Export start time in milliseconds
  TxMs1     : UDINT := 0;                        // Čas konca exportu v milisekundách ; Export end time in milliseconds
  TxDur     : UDINT := 0;                        // Trvanie exportu v milisekundách ; Export duration in milliseconds
  TxCyc     : UDINT := 0;                        // Počítadlo cyklov PLC ; PLC-cycle counter
  TxCyc0    : UDINT := 0;                        // Počítadlo cyklov pri štarte exportu ; PLC-cycle count at export start
  TxCycN    : UDINT := 0;                        // Počet cyklov spotrebovaných exportom ; Number of cycles used by the export
  TxDoneN   : UDINT := 0;                        // Počet dokončených viet ; Number of completed records
END_VAR

// Zapíše ľubovoľný úsek pamäte do otvoreného JSON súboru a kontroluje počet bajtov. ; Write a raw memory span to the open JSON file and verify the byte count.
FUNCTION TxWriteRaw : BOOL
  VAR_INPUT
    Pos : UDINT;  // Začiatočná adresa alebo offset zapisovaných dát ; Start address or offset of the data being written
    Siz : UDINT;  // Počet bajtov zapisovaného úseku ; Number of bytes in the section being written
  END_VAR
  VAR
    N : UDINT;  // Počet bajtov skutočne zapísaných funkciou ; Number of bytes actually written by the function
  END_VAR
  TxWriteRaw := FALSE;
  IF Siz = 0 THEN TxWriteRaw := TRUE; RETURN; END_IF;
  N := FileWrite(hFile := TxH, adrBuf := Pos, size := Siz);
  TxBytes := TxBytes + N;
  IF N <> Siz THEN TxWorkErr := 3; RETURN; END_IF;
  TxWriteRaw := TRUE;
END_FUNCTION

// Zapíše textový reťazec do exportného súboru. ; Write a text string to the export file.
FUNCTION TxWrite : BOOL
  VAR_INPUT
    Text : STRING[255];  // Textový obsah zapisovaný do JSON ; Text content being written to JSON
  END_VAR
  TxWrite := TxWriteRaw(Pos := PTR_TO_UDINT(ADR(Text)), Siz := INT_TO_UDINT(LEN(Text)));
END_FUNCTION

// Zapíše text medzi úvodzovky JSON. ; Write text enclosed in JSON quotes.
FUNCTION TxWriteQuoted : BOOL
  VAR_INPUT
    Text : STRING[255];  // Textový obsah zapisovaný do JSON ; Text content being written to JSON
  END_VAR
  TxWriteQuoted := FALSE;
  IF NOT TxWrite(Text := '"') THEN RETURN; END_IF;
  IF NOT TxWrite(Text := Text) THEN RETURN; END_IF;
  IF NOT TxWrite(Text := '"') THEN RETURN; END_IF;
  TxWriteQuoted := TRUE;
END_FUNCTION

// Prevedie reťazec PLC z CP1250 na UTF-8 a escapuje riadiace znaky JSON. ; Convert the PLC string from CP1250 to UTF-8 and escape JSON control characters.
// Prevedie PLC reťazec na korektný UTF-8 reťazec JSON. ; Convert a PLC string into valid UTF-8 JSON text.
// Skopíruje pevný úsek PLC STRING, prevedie CP1250 na UTF-8 a začne JSON reťazec. ; Copy a fixed PLC STRING span, convert CP1250 to UTF-8, and open a JSON string.
FUNCTION TxWriteString : BOOL
  VAR_INPUT
    Pos  : UDINT;  // Začiatočná adresa alebo offset zapisovaných dát ; Start address or offset of the data being written
    Span : UINT;   // Veľkosť hodnoty podľa schémy ; Value size from the schema
  END_VAR
  VAR
    Cp  : STRING[255];  // Počet bajtov v PLC reťazci ; Number of bytes in the PLC string
    Utf : STRING[255];  // Reťazec po prevode do UTF-8 ; String after conversion to UTF-8
    Src : PTR_TO BYTE;  // Ukazovateľ na zdrojové bajty ; Pointer to the source bytes
    P   : PTR_TO BYTE;  // Pracovný ukazovateľ na hodnotu ; Working pointer to the value
    H   : PTR_TO BYTE;  // Hexadecimálna číslica ; Hexadecimal digit
    Q   : PTR_TO BYTE;  // Pracovný znak pri escapovaní JSON ; Working character during JSON escaping
    B   : BYTE;         // Pracovný bajt hodnoty ; Working value byte
    N   : UDINT;        // Počet bajtov skutočne zapísaných funkciou ; Number of bytes actually written by the function
    I   : UINT;         // Index opakovania alebo poľa ; Loop or array index
    J   : UINT;         // Druhý index vnoreného prechodu ; Secondary index for nested traversal
  END_VAR
  TxWriteString := FALSE;
  IF (Span = 0) OR (Span > SIZEOF(Cp)) THEN TxWorkErr := 7; RETURN; END_IF;
  Cp := '';
  Utf := '';
  Src := UDINT_TO_PTR(Pos);
  N := MemCpyPtr(source := Src, dest := ADR(Cp), length := UINT_TO_UDINT(Span));
  IF N <> UINT_TO_UDINT(Span) THEN TxWorkErr := 7; RETURN; END_IF;
  N := CP1250_TO_UTF8(cp1250 := Cp, utf8 := Utf, maxLen := 255);
  IF (Cp <> '') AND (N = 0) THEN TxWorkErr := 7; RETURN; END_IF;
  IF NOT TxWrite(Text := '"') THEN RETURN; END_IF;
  P := ADR(Utf);
  H := ADR(TxHex);
  // Každý UTF-8 bajt zapíše priamo alebo ho escapuje podľa pravidiel JSON. ; Write each UTF-8 byte directly or escape it according to JSON rules.
  FOR I := 1 TO INT_TO_UINT(LEN(Utf)) DO
    B := P^;
    CASE B OF
      8:  IF NOT TxWrite(Text := '\b') THEN RETURN; END_IF;
      9:  IF NOT TxWrite(Text := '\t') THEN RETURN; END_IF;
      10: IF NOT TxWrite(Text := '\n') THEN RETURN; END_IF;
      12: IF NOT TxWrite(Text := '\f') THEN RETURN; END_IF;
      13: IF NOT TxWrite(Text := '\r') THEN RETURN; END_IF;
      34: IF NOT TxWrite(Text := '\"') THEN RETURN; END_IF;
      92: IF NOT TxWrite(Text := '\\') THEN RETURN; END_IF;
      ELSE
        IF B < 32 THEN
          IF NOT TxWrite(Text := '\u00') THEN RETURN; END_IF;
          Q := H;
          J := 0;
          WHILE J < BYTE_TO_UINT(B) / 16 DO Q := Q + 1; J := J + 1; END_WHILE;
          IF NOT TxWriteRaw(Pos := PTR_TO_UDINT(Q), Siz := 1) THEN RETURN; END_IF;
          Q := H;
          J := 0;
          WHILE J < BYTE_TO_UINT(B) MOD 16 DO Q := Q + 1; J := J + 1; END_WHILE;
          IF NOT TxWriteRaw(Pos := PTR_TO_UDINT(Q), Siz := 1) THEN RETURN; END_IF;
        ELSE
          IF NOT TxWriteRaw(Pos := PTR_TO_UDINT(P), Siz := 1) THEN RETURN; END_IF;
        END_IF;
    END_CASE;
    P := P + 1;
  END_FOR;
  IF NOT TxWrite(Text := '"') THEN RETURN; END_IF;
  TxWriteString := TRUE;
END_FUNCTION

// Načíta jednu hodnotu podľa typu v schéme a zapíše ju do JSON. ; Read one value according to its schema type and write it to JSON.
// Schéma dodá typ a adresu ; nižšie sa hodnota prečíta cez ukazovateľ správneho typu. ; The schema supplies type and address ; the value is read through a correctly typed pointer.
FUNCTION TxWriteValue : BOOL
  VAR_INPUT
    Parent : UDINT;  // Adresa rodičovskej štruktúry v mRam ; Address of the parent structure in mRam
    Nd     : UINT;   // Index uzla aktuálnej položky schémy ; Schema-node index of the current field
    El     : INT;    // Index prvku poľa ; Array element index
  END_VAR
  VAR
    ValAdr : UDINT;         // Adresa hodnoty v mRam ; Address of the value in mRam
    Tag    : USINT;         // Základný typ hodnoty ; Base type of the value
    BitPos : SINT;          // Pozícia BOOL v bajte ; BOOL bit position within its byte
    Mask   : UINT;          // Maska na vyčítanie jedného BOOL bitu ; Mask used to read one BOOL bit
    I      : SINT;          // Index opakovania alebo poľa ; Loop or array index
    Text   : STRING[255];   // Textový obsah zapisovaný do JSON ; Text content being written to JSON
    PB     : PTR_TO BYTE;
    PS     : PTR_TO SINT;
    PU     : PTR_TO USINT;
    PI     : PTR_TO INT;
    PUI    : PTR_TO UINT;
    PDI    : PTR_TO DINT;
    PUD    : PTR_TO UDINT;
    PW     : PTR_TO WORD;
    PDW    : PTR_TO DWORD;
    PR     : PTR_TO REAL;
    PLR    : PTR_TO LREAL;
    PT     : PTR_TO TIME;
    PDate  : PTR_TO DATE;
    PTod   : PTR_TO TOD;
    PDT    : PTR_TO DT;
  END_VAR
  TxWriteValue := FALSE;
  ValAdr := SchAdr(Parent := Parent, Nd := Nd, El := El);
  IF ValAdr = 0 THEN TxWorkErr := 6; RETURN; END_IF;
  Tag := aNode[Nd].Tag MOD SCH_ARRAY;

  // Vyberie prevod podľa IEC dátového typu položky. ; Select conversion according to the field's IEC data type.
  CASE Tag OF
    SCH_BOOL:
      PB := UDINT_TO_PTR(ValAdr);
      BitPos := SchBit(Nd := Nd, El := El);
      IF BitPos < 0 THEN TxWorkErr := 6; RETURN; END_IF;
      Mask := 1;
      FOR I := 1 TO BitPos DO Mask := Mask * 2; END_FOR;
      IF (BYTE_TO_UINT(PB^) / Mask) MOD 2 = 1 THEN Text := 'true'; ELSE Text := 'false'; END_IF;
    SCH_SINT: PS := UDINT_TO_PTR(ValAdr); Text := SINT_TO_STRING(PS^);
    SCH_USINT: PU := UDINT_TO_PTR(ValAdr); Text := USINT_TO_STRING(PU^);
    SCH_INT: PI := UDINT_TO_PTR(ValAdr); Text := INT_TO_STRING(PI^);
    SCH_UINT: PUI := UDINT_TO_PTR(ValAdr); Text := UINT_TO_STRING(PUI^);
    SCH_DINT: PDI := UDINT_TO_PTR(ValAdr); Text := DINT_TO_STRING(PDI^);
    SCH_UDINT: PUD := UDINT_TO_PTR(ValAdr); Text := UDINT_TO_STRING(PUD^);
    SCH_BYTE: PB := UDINT_TO_PTR(ValAdr); Text := UDINT_TO_STRING(BYTE_TO_UDINT(PB^));
    SCH_WORD: PW := UDINT_TO_PTR(ValAdr); Text := UDINT_TO_STRING(WORD_TO_UDINT(PW^));
    SCH_DWORD: PDW := UDINT_TO_PTR(ValAdr); Text := UDINT_TO_STRING(DWORD_TO_UDINT(PDW^));
    SCH_REAL: PR := UDINT_TO_PTR(ValAdr); Text := REAL_TO_STRING(PR^);
    SCH_LREAL: PLR := UDINT_TO_PTR(ValAdr); Text := LREAL_TO_STRING(PLR^);
    SCH_STRING:
      TxWriteValue := TxWriteString(Pos := ValAdr, Span := aNode[Nd].Span);
      RETURN;
    SCH_TIME: PT := UDINT_TO_PTR(ValAdr); Text := TIME_TO_STRING(PT^);
    SCH_DATE: PDate := UDINT_TO_PTR(ValAdr); Text := DATE_TO_STRING(PDate^);
    SCH_TIME_OF_DAY: PTod := UDINT_TO_PTR(ValAdr); Text := TOD_TO_STRING(PTod^);
    SCH_DATE_AND_TIME: PDT := UDINT_TO_PTR(ValAdr); Text := DT_TO_STRING(PDT^);
    ELSE TxWorkErr := 6; RETURN;
  END_CASE;

  IF (Tag = SCH_TIME) OR (Tag = SCH_DATE) OR (Tag = SCH_TIME_OF_DAY) OR (Tag = SCH_DATE_AND_TIME) THEN
    TxWriteValue := TxWriteQuoted(Text := Text);
  ELSE
    TxWriteValue := TxWrite(Text := Text);
  END_IF;
END_FUNCTION

// Prečíta PLC systémové hodiny v milisekundách pre meranie exportu. ; Read the PLC millisecond clock for export timing.
FUNCTION TxClockMs : UDINT
  VAR_EXTERNAL
    AT %SL52 : DWORD;
  END_VAR
  TxClockMs := DWORD_TO_UDINT(%SL52);
END_FUNCTION

// Zapíše jeden riadok do meracieho logu exportu. ; Write one line to the export measurement log.
FUNCTION TxLogPut : BOOL
  VAR_INPUT
    Hnd  : HANDLE;
    Text : STRING[255];  // Textový obsah zapisovaný do JSON ; Text content being written to JSON
  END_VAR
  VAR
    N : UDINT;  // Počet bajtov skutočne zapísaných funkciou ; Number of bytes actually written by the function
  END_VAR
  N := FileWrite(hFile := Hnd, adrBuf := PTR_TO_UDINT(ADR(Text)), size := INT_TO_UDINT(LEN(Text)));
  TxLogPut := N = INT_TO_UDINT(LEN(Text));
END_FUNCTION

// Zapíše parametre, výsledok a namerané trvanie exportu do tx.log. ; Write export parameters, result, and timing to tx.log.
FUNCTION TxWriteLog : BOOL
  VAR
    Hnd    : HANDLE;
    Line   : STRING[255];
    Closed : BOOL;          // Príznak úspešného uzatvorenia súboru ; Flag indicating the file closed successfully
    Ok     : BOOL := TRUE;  // Príznak úspešného zápisu ; Flag indicating a successful write
  END_VAR
  TxWriteLog := FALSE;
  Hnd := FileOpen(fileName := TxLogPath, mode := F_WRITE);
  IF Hnd = INVALID_HANDLE_VALUE THEN RETURN; END_IF;

  Line := CONCAT('api_V12 TX export', TxCRLF); Ok := Ok AND TxLogPut(Hnd := Hnd, Text := Line);
  Line := CONCAT('file=RAM/tx.json', TxCRLF); Ok := Ok AND TxLogPut(Hnd := Hnd, Text := Line);
  Line := CONCAT('rq=', UDINT_TO_STRING(TxRqW), TxCRLF); Ok := Ok AND TxLogPut(Hnd := Hnd, Text := Line);
  Line := CONCAT('cf=', USINT_TO_STRING(TxCfW), TxCRLF); Ok := Ok AND TxLogPut(Hnd := Hnd, Text := Line);
  IF (TxCfW >= 1) AND (TxCfW <= UINT_TO_USINT(SCH_DEF_N)) THEN
    Line := CONCAT('type=', aSch[TxCfW].Code, TxCRLF); Ok := Ok AND TxLogPut(Hnd := Hnd, Text := Line);
  END_IF;
  IF TxMode = 3 THEN Line := CONCAT('mode=all', TxCRLF);
  ELSIF TxMode = 2 THEN Line := CONCAT('mode=range', TxCRLF);
  ELSE Line := CONCAT('mode=one', TxCRLF);
  END_IF;
  Ok := Ok AND TxLogPut(Hnd := Hnd, Text := Line);
  Line := CONCAT('from=', UDINT_TO_STRING(TxFrom), TxCRLF); Ok := Ok AND TxLogPut(Hnd := Hnd, Text := Line);
  Line := CONCAT('to=', UDINT_TO_STRING(TxTo), TxCRLF); Ok := Ok AND TxLogPut(Hnd := Hnd, Text := Line);
  IF TxTo >= TxFrom THEN Line := CONCAT('records=', UDINT_TO_STRING(TxTo - TxFrom + 1), TxCRLF);
  ELSE Line := CONCAT('records=0', TxCRLF);
  END_IF;
  Ok := Ok AND TxLogPut(Hnd := Hnd, Text := Line);
  Line := CONCAT('records_done=', UDINT_TO_STRING(TxDoneN), TxCRLF); Ok := Ok AND TxLogPut(Hnd := Hnd, Text := Line);
  IF (TxCfW >= 1) AND (TxCfW <= UINT_TO_USINT(SCH_DEF_N)) THEN
    Line := CONCAT('record_bytes=', UDINT_TO_STRING(aSch[TxCfW].Siz), TxCRLF); Ok := Ok AND TxLogPut(Hnd := Hnd, Text := Line);
    Line := CONCAT('schema_nodes=', UINT_TO_STRING(aSch[TxCfW].Cnt), TxCRLF); Ok := Ok AND TxLogPut(Hnd := Hnd, Text := Line);
  END_IF;
  Line := CONCAT('json_bytes=', UDINT_TO_STRING(TxBytes), TxCRLF); Ok := Ok AND TxLogPut(Hnd := Hnd, Text := Line);
  Line := CONCAT('start_ms=', UDINT_TO_STRING(TxMs0), TxCRLF); Ok := Ok AND TxLogPut(Hnd := Hnd, Text := Line);
  Line := CONCAT('end_ms=', UDINT_TO_STRING(TxMs1), TxCRLF); Ok := Ok AND TxLogPut(Hnd := Hnd, Text := Line);
  Line := CONCAT('duration_ms=', UDINT_TO_STRING(TxDur), TxCRLF); Ok := Ok AND TxLogPut(Hnd := Hnd, Text := Line);
  Line := CONCAT('plc_cycles=', UDINT_TO_STRING(TxCycN), TxCRLF); Ok := Ok AND TxLogPut(Hnd := Hnd, Text := Line);
  IF TxWorkErr = 0 THEN Line := CONCAT('result=OK', TxCRLF);
  ELSE Line := CONCAT('result=ERROR', TxCRLF);
  END_IF;
  Ok := Ok AND TxLogPut(Hnd := Hnd, Text := Line);
  Line := CONCAT('error=', USINT_TO_STRING(TxWorkErr), TxCRLF); Ok := Ok AND TxLogPut(Hnd := Hnd, Text := Line);

  Closed := FileClose(hFile := Hnd);
  TxWriteLog := Ok AND Closed;
END_FUNCTION

// Prejde uzly jednej vety podľa schémy a vytvorí jej vnorený JSON objekt. ; Traverse one record's schema nodes and produce its nested JSON object.
// Zásobníky Kind/Base/StartNd/EndNd riadia iteratívny prechod vnorenými objektmi a poľami STRUCT. ; Kind/Base/StartNd/EndNd stacks drive iterative traversal of nested STRUCT objects and arrays.
FUNCTION TxWriteRecord : BOOL
  VAR_INPUT
    Cf  : USINT;  // Index typu vybraného pre operáciu ; Index of the type selected for the operation
    Rec : UDINT;  // Číslo spracúvanej vety ; Number of the record being processed
  END_VAR
  VAR
    Root    : UDINT;                  // Adresa koreňa vybranej vety ; Root address of the selected record
    Nd      : UINT;                   // Index uzla aktuálnej položky schémy ; Schema-node index of the current field
    NextNd  : UINT;                   // Index nasledujúceho uzla schémy ; Index of the next schema node
    Tag     : USINT;                  // Základný typ hodnoty ; Base type of the value
    D       : INT;                    // Hĺbka zásobníka vnorených objektov ; Nested-object stack depth
    ElNow   : INT;
    ElLast  : INT;
    Head    : STRING[40];             // Názov JSON poľa vrátane dvojbodky ; JSON field name including its colon
    Done    : BOOL;                   // Príznak dokončenia aktuálnej vety ; Flag indicating the current record is complete
    Kind    : ARRAY[0..15] OF USINT;  // Typ rámca v zásobníku prechodu ; Frame kind in the traversal stack ; 1=object, 2=array-of-struct controller
    Base    : ARRAY[0..15] OF UDINT;  // Základná adresa rámca v mRam ; Base address of the frame in mRam
    First   : ARRAY[0..15] OF BOOL;   // Prvý uzol aktuálneho objektu ; First node of the current object
    StartNd : ARRAY[0..15] OF UINT;   // Prvý uzol potomkov aktuálneho objektu ; First child node of the current object
    EndNd   : ARRAY[0..15] OF UINT;   // Koniec rozsahu uzlov aktuálneho objektu ; End of the current object's node range
    AfterNd : ARRAY[0..15] OF UINT;   // Prvý uzol nasledujúci po objekte ; First node after the object
    ArrNd   : ARRAY[0..15] OF UINT;   // Uzol poľa spracúvaný daným rámcom ; Array node processed by this frame
    ArrEl   : ARRAY[0..15] OF INT;    // Aktuálny IEC index prvku poľa ; Current IEC array element index
    ArrLast : ARRAY[0..15] OF INT;    // Posledný IEC index prvku poľa ; Last IEC array element index
  END_VAR

  TxWriteRecord := FALSE;
  Root := SchRoot(Cf := Cf, Rec := Rec);
  IF Root = 0 THEN TxWorkErr := 1; RETURN; END_IF;
  IF NOT TxWrite(Text := '{') THEN RETURN; END_IF;

  D := 0;
  Kind[0] := 1;
  Base[0] := Root;
  First[0] := TRUE;
  StartNd[0] := aSch[Cf].Fst;
  EndNd[0] := aSch[Cf].Fst + aSch[Cf].Cnt;
  Nd := StartNd[0];

  // Pokračuje, kým sa neuzavrie koreňový objekt alebo nevznikne chyba. ; Continue until the root object closes or an error occurs.
  WHILE NOT Done AND (TxWorkErr = 0) DO
    // Kontrola chráni stavový automat pred neplatným typom rámca zásobníka. ; Guard the state machine against an invalid stack-frame kind.
    IF Kind[D] <> 1 THEN TxWorkErr := 8;
    ELSIF Nd >= EndNd[D] THEN
      IF NOT TxWrite(Text := '}') THEN RETURN; END_IF;
      IF D = 0 THEN
        Done := TRUE;
      ELSE
        NextNd := AfterNd[D];
        D := D - 1;
        IF Kind[D] = 2 THEN
          IF ArrEl[D] < ArrLast[D] THEN
            ArrEl[D] := ArrEl[D] + 1;
            IF NOT TxWrite(Text := ',{') THEN RETURN; END_IF;
            IF D >= 15 THEN TxWorkErr := 5; RETURN; END_IF;
            D := D + 1;
            Kind[D] := 1;
            Base[D] := SchAdr(Parent := Base[D - 1], Nd := ArrNd[D - 1], El := ArrEl[D - 1]);
            First[D] := TRUE;
            StartNd[D] := StartNd[D - 1];
            EndNd[D] := EndNd[D - 1];
            AfterNd[D] := EndNd[D];
            Nd := StartNd[D];
          ELSE
            IF NOT TxWrite(Text := ']') THEN RETURN; END_IF;
            NextNd := AfterNd[D];
            D := D - 1;
            Nd := NextNd;
          END_IF;
        ELSE
          Nd := NextNd;
        END_IF;
      END_IF;
    ELSE
      IF NOT First[D] THEN IF NOT TxWrite(Text := ',') THEN RETURN; END_IF; END_IF;
      Head := CONCAT('"', aNode[Nd].Nam, '":');
      IF NOT TxWrite(Text := Head) THEN RETURN; END_IF;
      First[D] := FALSE;
      Tag := aNode[Nd].Tag MOD SCH_ARRAY;

      // Vnorený objekt alebo pole štruktúr sa spracuje rekurzívne simulovaným zásobníkom. ; Nested objects and STRUCT arrays are traversed with an explicit stack.
      IF Tag = SCH_STRUCT THEN
        NextNd := Nd + 1 + aNode[Nd].Aux;
        IF aNode[Nd].Tag >= SCH_ARRAY THEN
          IF (aNode[Nd].Cnt = 0) OR (D > 13) THEN TxWorkErr := 5; RETURN; END_IF;
          IF NOT TxWrite(Text := '[{') THEN RETURN; END_IF;
          D := D + 1;
          Kind[D] := 2;
          Base[D] := Base[D - 1];
          StartNd[D] := Nd + 1;
          EndNd[D] := NextNd;
          AfterNd[D] := NextNd;
          ArrNd[D] := Nd;
          ArrEl[D] := aNode[Nd].Lo;
          ArrLast[D] := aNode[Nd].Lo + UINT_TO_INT(aNode[Nd].Cnt) - 1;
          D := D + 1;
          Kind[D] := 1;
          Base[D] := SchAdr(Parent := Base[D - 1], Nd := ArrNd[D - 1], El := ArrEl[D - 1]);
          First[D] := TRUE;
          StartNd[D] := StartNd[D - 1];
          EndNd[D] := EndNd[D - 1];
          AfterNd[D] := EndNd[D];
          Nd := StartNd[D];
        ELSE
          IF D >= 15 THEN TxWorkErr := 5; RETURN; END_IF;
          IF NOT TxWrite(Text := '{') THEN RETURN; END_IF;
          D := D + 1;
          Kind[D] := 1;
          Base[D] := SchAdr(Parent := Base[D - 1], Nd := Nd, El := 0);
          First[D] := TRUE;
          StartNd[D] := Nd + 1;
          EndNd[D] := NextNd;
          AfterNd[D] := NextNd;
          Nd := StartNd[D];
        END_IF;
      ELSE
        IF aNode[Nd].Tag >= SCH_ARRAY THEN
          IF NOT TxWrite(Text := '[') THEN RETURN; END_IF;
          ElNow := aNode[Nd].Lo;
          ElLast := aNode[Nd].Lo + UINT_TO_INT(aNode[Nd].Cnt) - 1;
          WHILE (ElNow <= ElLast) AND (TxWorkErr = 0) DO
            IF ElNow > aNode[Nd].Lo THEN IF NOT TxWrite(Text := ',') THEN RETURN; END_IF; END_IF;
            IF NOT TxWriteValue(Parent := Base[D], Nd := Nd, El := ElNow) THEN RETURN; END_IF;
            ElNow := ElNow + 1;
          END_WHILE;
          IF NOT TxWrite(Text := ']') THEN RETURN; END_IF;
        ELSE
          IF NOT TxWriteValue(Parent := Base[D], Nd := Nd, El := 0) THEN RETURN; END_IF;
        END_IF;
        Nd := Nd + 1;
      END_IF;
    END_IF;
  END_WHILE;

  IF NOT Done AND (TxWorkErr = 0) THEN TxWorkErr := 8; END_IF;
  TxWriteRecord := Done AND (TxWorkErr = 0);
END_FUNCTION

// Uzatvorí export, zapíše log a potvrdí požiadavku klientovi. ; Close the export, write its log, and acknowledge the client request.
FUNCTION TxEnd : BOOL
  VAR
    Closed : BOOL := TRUE;  // Príznak úspešného uzatvorenia súboru ; Flag indicating the file closed successfully
    LogOk  : BOOL;          // Výsledok zápisu meracieho logu ; Result of writing the measurement log
  END_VAR
  IF TxH <> INVALID_HANDLE_VALUE THEN Closed := FileClose(hFile := TxH); END_IF;
  TxH := INVALID_HANDLE_VALUE;
  IF (TxWorkErr = 0) AND NOT Closed THEN TxWorkErr := 4; END_IF;
  TxMs1 := TxClockMs();
  TxDur := TxMs1 - TxMs0;
  TxCycN := TxCyc - TxCyc0 + 1;
  LogOk := TxWriteLog();
  IF (TxWorkErr = 0) AND NOT LogOk THEN TxWorkErr := 9; END_IF;
  TxErr := TxWorkErr;
  TxDone := TxRqW;
  TxSt := 0;
  TxEnd := TxWorkErr = 0;
END_FUNCTION

// Overí požiadavku, otvorí tx.json a zapíše hlavičku JSON obálky. ; Validate the request, open tx.json, and write the JSON envelope header.
// Overí požiadavku a pripraví export jednej alebo všetkých viet daného typu. ; Validate the request and prepare an export of one or all records of the selected type.
FUNCTION TxStart : BOOL
  VAR_INPUT
    Cf  : USINT;  // Index typu vybraného pre operáciu ; Index of the type selected for the operation
    Rec : UDINT;  // Číslo spracúvanej vety ; Number of the record being processed
    Rq  : UDINT;  // Číslo požiadavky klienta ; Client request number
  END_VAR
  VAR
    Ok : BOOL;  // Príznak úspešného zápisu ; Flag indicating a successful write
  END_VAR
  TxStart := FALSE;
  TxCfW := Cf;
  TxRqW := Rq;
  TxFrom := 0;
  TxTo := 0;
  TxNow := 0;
  TxMode := 0;
  TxDoneN := 0;
  TxBytes := 0;
  TxWorkErr := 0;
  TxMs0 := TxClockMs();
  TxCyc0 := TxCyc;
  TxErr := 1;

  IF NOT SchInit() OR (Cf < 1) OR (Cf > UINT_TO_USINT(SCH_DEF_N)) THEN
    TxWorkErr := 1; Ok := TxEnd(); RETURN;
  END_IF;
  // Nula vyberá všetky vety typu ; inak sa exportuje zadané číslo. ; Zero selects all records of the type ; otherwise export the requested record.
  IF Rec = 0 THEN
    TxMode := 3;
    TxFrom := 1;
    TxTo := aCfg[Cf].Rec;
  ELSE
    TxMode := 1;
    TxFrom := Rec;
    TxTo := Rec;
  END_IF;
  TxNow := TxFrom;
  IF (TxFrom < 1) OR (TxTo < TxFrom) OR (TxTo > aCfg[Cf].Rec) OR
     (SchRoot(Cf := Cf, Rec := TxFrom) = 0) OR (SchRoot(Cf := Cf, Rec := TxTo) = 0) THEN
    TxWorkErr := 1; Ok := TxEnd(); RETURN;
  END_IF;

  TxH := FileOpen(fileName := TxPath, mode := F_WRITE);
  IF TxH = INVALID_HANDLE_VALUE THEN TxWorkErr := 2; Ok := TxEnd(); RETURN; END_IF;

  // Zapíše hlavičku obálky s identifikátorom požiadavky a neskôr doplní rozsah i dáta. ; Write the request envelope header, then append range metadata and data.
  IF NOT TxWrite(Text := '{"rq":') THEN Ok := TxEnd(); RETURN; END_IF;
  IF NOT TxWrite(Text := UDINT_TO_STRING(Rq)) THEN Ok := TxEnd(); RETURN; END_IF;
  IF NOT TxWrite(Text := ',"cf":') THEN Ok := TxEnd(); RETURN; END_IF;
  IF NOT TxWrite(Text := USINT_TO_STRING(Cf)) THEN Ok := TxEnd(); RETURN; END_IF;
  IF NOT TxWrite(Text := ',"type":"') THEN Ok := TxEnd(); RETURN; END_IF;
  IF NOT TxWrite(Text := aSch[Cf].Code) THEN Ok := TxEnd(); RETURN; END_IF;
  IF NOT TxWrite(Text := '","from":') THEN Ok := TxEnd(); RETURN; END_IF;
  IF NOT TxWrite(Text := UDINT_TO_STRING(TxFrom)) THEN Ok := TxEnd(); RETURN; END_IF;
  IF NOT TxWrite(Text := ',"to":') THEN Ok := TxEnd(); RETURN; END_IF;
  IF NOT TxWrite(Text := UDINT_TO_STRING(TxTo)) THEN Ok := TxEnd(); RETURN; END_IF;
  IF NOT TxWrite(Text := ',"count":') THEN Ok := TxEnd(); RETURN; END_IF;
  IF NOT TxWrite(Text := UDINT_TO_STRING(TxTo - TxFrom + 1)) THEN Ok := TxEnd(); RETURN; END_IF;
  IF NOT TxWrite(Text := ',"data":[') THEN Ok := TxEnd(); RETURN; END_IF;
  TxSt := 1;
  TxStart := TRUE;
END_FUNCTION

// Stavový automat exportu ; na cyklus PLC spracuje najviac jednu vetu. ; Export state machine ; processes at most one record per PLC cycle.
// Nové TxRq založí export ; ďalšie cykly postupne dopíšu záznamy. ; A new TxRq starts an export ; subsequent cycles append records.
FUNCTION TxCycle : BOOL
  VAR
    Ok : BOOL;  // Príznak úspešného zápisu ; Flag indicating a successful write
  END_VAR
  TxCyc := TxCyc + 1;
  TxCycle := TRUE;

  // V nečinnom stave čaká na nové číslo požiadavky. ; While idle, wait for a new request number.
  IF TxSt = 0 THEN
    IF (TxRq = 0) OR (TxRq = TxSeen) THEN RETURN; END_IF;
    TxSeen := TxRq;
    TxCycle := TxStart(Cf := TxCf, Rec := TxRec, Rq := TxRq);
    RETURN;
  END_IF;

  IF TxSt <> 1 THEN TxWorkErr := 8; TxCycle := TxEnd(); RETURN; END_IF;
  // Ochrana pred prekročením koncového čísla vybraného rozsahu. ; Guard against passing the selected range's final record.
  IF TxNow > TxTo THEN TxWorkErr := 8; TxCycle := TxEnd(); RETURN; END_IF;

  IF TxNow > TxFrom THEN IF NOT TxWrite(Text := ',') THEN TxCycle := TxEnd(); RETURN; END_IF; END_IF;
  IF NOT TxWrite(Text := '{"rec":') THEN TxCycle := TxEnd(); RETURN; END_IF;
  IF NOT TxWrite(Text := UDINT_TO_STRING(TxNow)) THEN TxCycle := TxEnd(); RETURN; END_IF;
  IF NOT TxWrite(Text := ',"value":') THEN TxCycle := TxEnd(); RETURN; END_IF;
  IF NOT TxWriteRecord(Cf := TxCfW, Rec := TxNow) THEN TxCycle := TxEnd(); RETURN; END_IF;
  IF NOT TxWrite(Text := '}') THEN TxCycle := TxEnd(); RETURN; END_IF;
  TxDoneN := TxDoneN + 1;
  TxNow := TxNow + 1;

  IF TxNow > TxTo THEN
    IF NOT TxWrite(Text := ']}') THEN TxCycle := TxEnd(); RETURN; END_IF;
    Ok := TxEnd();
    TxCycle := Ok;
  END_IF;
END_FUNCTION

(* ---- _06_RxJson.ST ---- *)
VAR_GLOBAL
  RxPath        : STRING[80] := '//RAM/rx.json';  // Zdrojový súbor prijatého JSON ; Source file containing received JSON
  RxLogPath     : STRING[80] := '//RAM/rx.log';   // Súbor meraní importu ; Import measurement log file
  RxParser      : fbJsonFileParser;               // Parser súborového JSON ; File-based JSON parser
  RxInfo        : TJsonInfo;                      // Aktuálna položka vrátená parserom ; Current item returned by the parser
  RxTmp         : ARRAY[0.._NH_RAM] OF BYTE;      // Pracovná kópia dát pred potvrdením do mRam ; Staging copy before committing data to mRam
  RxLeafSeen    : ARRAY[1..SCH_LEAF_N] OF BOOL;   // Príznaky už načítaných povinných polí ; Flags for required fields already read
  RxSt          : USINT := 0;                     // Stavový automat importu ; Import state-machine state
  RxRqSeen      : UDINT := 0;                     // Posledná požiadavka už spracovaná PLC ; Latest request already processed by the PLC
  RxRqW         : UDINT := 0;                     // Číslo práve spracúvanej požiadavky ; Request number currently being processed
  RxWorkErr     : USINT := 0;                     // Pracovný kód chyby importu ; Working import error code
  RxErrTxt      : STRING[80] := '';               // Textový opis poslednej chyby ; Text description of the latest error
  RxLastName    : STRING[255] := '';              // Názov poslednej položky JSON ; Name of the latest JSON item
  RxCfW         : USINT := 0;                     // Typ vybraný pre aktuálny import ; Type selected for the current import
  RxTypeW       : STRING[4] := '';                // Kód typu uvedený v obálke JSON ; Type code supplied in the JSON envelope
  RxFrom        : UDINT := 0;                     // Prvá importovaná veta ; First record to import
  RxTo          : UDINT := 0;                     // Posledná importovaná veta ; Last record to import
  RxCount       : UDINT := 0;                     // Očakávaný počet importovaných viet ; Expected number of imported records
  RxFileRq      : UDINT := 0;                     // Číslo požiadavky zapísané v JSON ; Request number stored in the JSON file
  RxHdrCf       : BOOL := FALSE;                  // Príznak načítania typu v obálke ; Flag indicating the type was read from the envelope
  RxHdrType     : BOOL := FALSE;                  // Príznak načítania kódu typu ; Flag indicating the type code was read
  RxHdrFrom     : BOOL := FALSE;                  // Príznak načítania začiatku rozsahu ; Flag indicating the range start was read
  RxHdrTo       : BOOL := FALSE;                  // Príznak načítania konca rozsahu ; Flag indicating the range end was read
  RxHdrCount    : BOOL := FALSE;                  // Príznak načítania počtu viet ; Flag indicating the record count was read
  RxPrepared    : BOOL := FALSE;                  // TRUE po príprave pracovnej kópie ; TRUE after the staging copy is prepared
  RxHaveRec     : BOOL := FALSE;                  // TRUE, keď sa práve spracúva veta ; TRUE while a record is being processed
  RxIdx         : UINT := 0;                      // Index aktuálnej položky parsera ; Index of the current parser item
  RxRecCur      : UDINT := 0;                     // Číslo práve spracúvanej vety ; Number of the record currently being processed
  RxFieldsCur   : UINT := 0;                      // Počet polí načítaných v aktuálnej vete ; Fields read in the current record
  RxFieldsDone  : UDINT := 0;                     // Celkový počet úspešne načítaných polí ; Total number of fields read successfully
  RxRecordsDone : UDINT := 0;                     // Celkový počet úspešne načítaných viet ; Total number of records read successfully
  RxStageBytes  : UDINT := 0;                     // Veľkosť pracovnej kópie v bajtoch ; Staging-copy size in bytes
  RxMs0         : UDINT := 0;                     // Čas začiatku importu v milisekundách ; Import start time in milliseconds
  RxMs1         : UDINT := 0;                     // Čas konca importu v milisekundách ; Import end time in milliseconds
  RxDur         : UDINT := 0;                     // Trvanie importu v milisekundách ; Import duration in milliseconds
  RxCyc         : UDINT := 0;                     // Počítadlo cyklov PLC ; PLC-cycle counter
  RxCyc0        : UDINT := 0;                     // Počítadlo cyklov pri štarte importu ; PLC-cycle count at import start
  RxCycN        : UDINT := 0;                     // Počet cyklov spotrebovaných importom ; Number of cycles used by the import
  RxCommitted   : BOOL := FALSE;
END_VAR

// Po načítaní hlavičky pripraví kópiu záznamov v pomocnej pamäti. ; Prepare a record copy in staging memory after reading the envelope.
// Overí hlavičku a rozsah a skopíruje pôvodné vety do pomocnej pamäte. ; Validate the header and range, then copy the existing records to staging memory.
// Validuje identitu typu, číslovanie viet a veľkosť staging priestoru ešte pred zmenou dát. ; Validate type identity, record numbering, and staging capacity before changing data.
FUNCTION RxPrepare : BOOL
  VAR
    Copied : UDINT;  // Počet bajtov skopírovaných do pracovnej pamäte ; Number of bytes copied to staging memory
  END_VAR
  RxPrepare := FALSE;
  IF RxPrepared THEN RxPrepare := TRUE; RETURN; END_IF;
  IF NOT RxHdrCf OR NOT RxHdrType OR NOT RxHdrFrom OR NOT RxHdrTo OR NOT RxHdrCount THEN
    RxWorkErr := 3; RxErrTxt := 'Incomplete header'; RETURN;
  END_IF;
  IF RxFileRq <> RxRqW THEN
    RxWorkErr := 3; RxErrTxt := 'Request number mismatch'; RETURN;
  END_IF;
  IF (RxCfW < 1) OR (RxCfW > UINT_TO_USINT(SCH_DEF_N)) THEN
    RxWorkErr := 3; RxErrTxt := 'Invalid cf'; RETURN;
  END_IF;
  IF RxTypeW <> aSch[RxCfW].Code THEN
    RxWorkErr := 3; RxErrTxt := 'Type does not match cf'; RETURN;
  END_IF;
  IF (RxFrom < 1) OR (RxTo < RxFrom) OR (RxTo > aCfg[RxCfW].Rec) OR
     (RxCount <> RxTo - RxFrom + 1) THEN
    RxWorkErr := 3; RxErrTxt := 'Invalid record range'; RETURN;
  END_IF;
  RxStageBytes := RxCount * aSch[RxCfW].Siz;
  IF (RxStageBytes = 0) OR (RxStageBytes > SIZEOF(RxTmp)) THEN
    RxWorkErr := 3; RxErrTxt := 'Staging buffer too small'; RETURN;
  END_IF;
  Copied := MemCpyPtr(  // Vytvorí pracovnú kópiu pôvodného rozsahu ; neúplný alebo chybný JSON tak nemení mRam. ; Create a working copy of the original range so incomplete or invalid JSON cannot alter mRam.
    source := UDINT_TO_PTR(aCfg[RxCfW].Ram + (RxFrom - 1) * aSch[RxCfW].Siz),
    dest := ADR(RxTmp[0]), length := RxStageBytes);
  IF Copied <> RxStageBytes THEN RxWorkErr := 7; RxErrTxt := 'Staging copy failed'; RETURN; END_IF;
  RxPrepared := TRUE;
  RxPrepare := TRUE;
END_FUNCTION

// Prevedie jednu hodnotu JSON na PLC typ a uloží ju do pomocnej pamäte. ; Convert one JSON value to its PLC type and store it in staging memory.
// Prevedie skalárnu hodnotu JSON na typ a rozloženie určené schémou. ; Convert a JSON scalar to the type and layout specified by the schema.
// Každý typ sa prevedie oddelene ; BOOL mení iba príslušný bit a STRING sa konvertuje do CP1250. ; Convert each type explicitly ; BOOL updates one bit and STRING is converted to CP1250.
FUNCTION RxSetValue : BOOL
  VAR_INPUT
    Lf    : UINT;         // Index cieľového poľa v schéme ; Target leaf-field index in the schema
    Pos   : UDINT;        // Adresa alebo pozícia hodnoty v pracovnej pamäti ; Address or position of the value in staging memory
    Value : STRING[255];  // Hodnota načítaná z JSON parsera ; Value read from the JSON parser
  END_VAR
  VAR
    Tmp    : STRING[255];   // Pracovná hodnota počas typovej konverzie ; Temporary value during type conversion
    N      : UDINT;         // Počet bajtov skopírovaných alebo zapísaných ; Number of bytes copied or written
    U      : UINT;          // Medzivýsledok prevodu na celé číslo bez znamienka ; Intermediate unsigned-integer conversion value
    Mask   : UINT;          // Maska pre nastavenie alebo kontrolu bitu ; Mask used to set or check a bit
    I      : SINT;          // Index bajtu alebo prvku poľa ; Byte or array-element index
    BitMax : SINT;          // Počet platných bitov poľa BOOL ; Number of valid BOOL-array bits
    PB     : PTR_TO BYTE;   // Ukazovateľ na bajt cieľovej hodnoty ; Pointer to a byte of the target value
    PS     : PTR_TO SINT;   // Ukazovateľ na hodnotu typu SINT ; Pointer to a SINT value
    PU     : PTR_TO USINT;  // Ukazovateľ na hodnotu typu USINT ; Pointer to a USINT value
    PI     : PTR_TO INT;    // Ukazovateľ na hodnotu typu INT ; Pointer to an INT value
    PUI    : PTR_TO UINT;   // Ukazovateľ na hodnotu typu UINT ; Pointer to a UINT value
    PDI    : PTR_TO DINT;   // Ukazovateľ na hodnotu typu DINT ; Pointer to a DINT value
    PUD    : PTR_TO UDINT;  // Ukazovateľ na hodnotu typu UDINT ; Pointer to a UDINT value
    PW     : PTR_TO WORD;   // Ukazovateľ na hodnotu typu WORD ; Pointer to a WORD value
    PDW    : PTR_TO DWORD;  // Ukazovateľ na hodnotu typu DWORD ; Pointer to a DWORD value
    PR     : PTR_TO REAL;   // Ukazovateľ na hodnotu typu REAL ; Pointer to a REAL value
    PLR    : PTR_TO LREAL;  // Ukazovateľ na hodnotu typu LREAL ; Pointer to an LREAL value
    PT     : PTR_TO TIME;   // Ukazovateľ na hodnotu typu TIME ; Pointer to a TIME value
    PDate  : PTR_TO DATE;   // Ukazovateľ na hodnotu typu DATE ; Pointer to a DATE value
    PTod   : PTR_TO TOD;    // Ukazovateľ na hodnotu typu TOD ; Pointer to a TOD value
    PDT    : PTR_TO DT;     // Ukazovateľ na hodnotu typu DT ; Pointer to a DT value
  END_VAR
  RxSetValue := FALSE;
  IF (Lf < 1) OR (Lf > SCH_LEAF_N) OR (Pos = 0) THEN
    RxWorkErr := 6; RxErrTxt := 'Invalid leaf address'; RETURN;
  END_IF;
  Tmp := Value;
  PB := UDINT_TO_PTR(Pos);
  // Konverzia vychádza z typu poľa v tabuľke schémy, nie z odhadu klienta. ; Conversion uses the field type from the schema table, not a client-side guess.
  CASE aLeaf[Lf].Tag OF
    SCH_BOOL:
      IF (Tmp <> 'true') AND (Tmp <> 'false') AND (Tmp <> '1') AND (Tmp <> '0') THEN
        RxWorkErr := 6; RxErrTxt := 'Invalid BOOL'; RETURN;
      END_IF;
      Mask := 1;
      BitMax := aLeaf[Lf].BitPos;
      FOR I := 1 TO BitMax DO Mask := Mask * 2; END_FOR;
      U := BYTE_TO_UINT(PB^);
      IF (Tmp = 'true') OR (Tmp = '1') THEN
        IF (U / Mask) MOD 2 = 0 THEN PB^ := UDINT_TO_BYTE(UINT_TO_UDINT(U + Mask)); END_IF;
      ELSE
        IF (U / Mask) MOD 2 = 1 THEN PB^ := UDINT_TO_BYTE(UINT_TO_UDINT(U - Mask)); END_IF;
      END_IF;
    SCH_SINT: PS := UDINT_TO_PTR(Pos); PS^ := STRING_TO_SINT(Tmp);
    SCH_USINT: PU := UDINT_TO_PTR(Pos); PU^ := STRING_TO_USINT(Tmp);
    SCH_INT: PI := UDINT_TO_PTR(Pos); PI^ := STRING_TO_INT(Tmp);
    SCH_UINT: PUI := UDINT_TO_PTR(Pos); PUI^ := STRING_TO_UINT(Tmp);
    SCH_DINT: PDI := UDINT_TO_PTR(Pos); PDI^ := STRING_TO_DINT(Tmp);
    SCH_UDINT: PUD := UDINT_TO_PTR(Pos); PUD^ := STRING_TO_UDINT(Tmp);
    SCH_BYTE: PB := UDINT_TO_PTR(Pos); PB^ := UDINT_TO_BYTE(STRING_TO_UDINT(Tmp));
    SCH_WORD: PW := UDINT_TO_PTR(Pos); PW^ := UDINT_TO_WORD(STRING_TO_UDINT(Tmp));
    SCH_DWORD: PDW := UDINT_TO_PTR(Pos); PDW^ := UDINT_TO_DWORD(STRING_TO_UDINT(Tmp));
    SCH_REAL: PR := UDINT_TO_PTR(Pos); PR^ := STRING_TO_REAL_EX(Tmp);
    SCH_LREAL: PLR := UDINT_TO_PTR(Pos); PLR^ := STRING_TO_LREAL_EX(Tmp);
    SCH_STRING:
      U := UTF8_TO_CP125x(str := Tmp, codePage := 1250);
      IF UINT_TO_UDINT(U) >= UINT_TO_UDINT(aLeaf[Lf].Span) THEN
        RxWorkErr := 6; RxErrTxt := 'STRING too long'; RETURN;
      END_IF;
      MemsetPtr(dest := PB, val := 0, length := aLeaf[Lf].Span);
      N := MemCpyPtr(source := ADR(Tmp), dest := PB, length := UINT_TO_UDINT(U) + 1);
      IF N <> UINT_TO_UDINT(U) + 1 THEN RxWorkErr := 6; RxErrTxt := 'STRING copy failed'; RETURN; END_IF;
    SCH_TIME: PT := UDINT_TO_PTR(Pos); PT^ := STRING_TO_TIME(Tmp);
    SCH_DATE: PDate := UDINT_TO_PTR(Pos); PDate^ := STRING_TO_DATE(Tmp);
    SCH_TIME_OF_DAY: PTod := UDINT_TO_PTR(Pos); PTod^ := STRING_TO_TOD(Tmp);
    SCH_DATE_AND_TIME: PDT := UDINT_TO_PTR(Pos); PDT^ := STRING_TO_DT(Tmp);
    ELSE RxWorkErr := 6; RxErrTxt := 'Unsupported type'; RETURN;
  END_CASE;
  RxSetValue := TRUE;
END_FUNCTION

// Zapíše priebeh, počty polí, chybu a čas importu do rx.log. ; Write import progress, field counts, errors, and timing to rx.log.
FUNCTION RxWriteLog : BOOL
  VAR
    Hnd    : HANDLE;        // Handle otvoreného súboru logu ; Handle of the open log file
    Line   : STRING[255];   // Pripravovaný riadok logu ; Log line being prepared
    Closed : BOOL;          // Výsledok uzatvorenia súboru ; Result of closing the file
    Ok     : BOOL := TRUE;  // Príznak úspešného dokončenia kroku ; Flag indicating the step completed successfully
  END_VAR
  RxWriteLog := FALSE;
  Hnd := FileOpen(fileName := RxLogPath, mode := F_WRITE);
  IF Hnd = INVALID_HANDLE_VALUE THEN RETURN; END_IF;
  Line := CONCAT('api_V12 RX import', TxCRLF); Ok := Ok AND TxLogPut(Hnd := Hnd, Text := Line);
  Line := CONCAT('file=RAM/rx.json', TxCRLF); Ok := Ok AND TxLogPut(Hnd := Hnd, Text := Line);
  Line := CONCAT('request=', UDINT_TO_STRING(RxRqW), TxCRLF); Ok := Ok AND TxLogPut(Hnd := Hnd, Text := Line);
  Line := CONCAT('file_rq=', UDINT_TO_STRING(RxFileRq), TxCRLF); Ok := Ok AND TxLogPut(Hnd := Hnd, Text := Line);
  Line := CONCAT('cf=', USINT_TO_STRING(RxCfW), TxCRLF); Ok := Ok AND TxLogPut(Hnd := Hnd, Text := Line);
  Line := CONCAT('type=', RxTypeW, TxCRLF); Ok := Ok AND TxLogPut(Hnd := Hnd, Text := Line);
  Line := CONCAT('from=', UDINT_TO_STRING(RxFrom), TxCRLF); Ok := Ok AND TxLogPut(Hnd := Hnd, Text := Line);
  Line := CONCAT('to=', UDINT_TO_STRING(RxTo), TxCRLF); Ok := Ok AND TxLogPut(Hnd := Hnd, Text := Line);
  Line := CONCAT('records=', UDINT_TO_STRING(RxCount), TxCRLF); Ok := Ok AND TxLogPut(Hnd := Hnd, Text := Line);
  Line := CONCAT('records_done=', UDINT_TO_STRING(RxRecordsDone), TxCRLF); Ok := Ok AND TxLogPut(Hnd := Hnd, Text := Line);
  Line := CONCAT('fields_done=', UDINT_TO_STRING(RxFieldsDone), TxCRLF); Ok := Ok AND TxLogPut(Hnd := Hnd, Text := Line);
  Line := CONCAT('file_bytes=', UDINT_TO_STRING(RxParser.fileSize), TxCRLF); Ok := Ok AND TxLogPut(Hnd := Hnd, Text := Line);
  Line := CONCAT('processed_bytes=', UDINT_TO_STRING(RxParser.processed), TxCRLF); Ok := Ok AND TxLogPut(Hnd := Hnd, Text := Line);
  Line := CONCAT('last_item=', RxLastName, TxCRLF); Ok := Ok AND TxLogPut(Hnd := Hnd, Text := Line);
  Line := CONCAT('staged_bytes=', UDINT_TO_STRING(RxStageBytes), TxCRLF); Ok := Ok AND TxLogPut(Hnd := Hnd, Text := Line);
  Line := CONCAT('start_ms=', UDINT_TO_STRING(RxMs0), TxCRLF); Ok := Ok AND TxLogPut(Hnd := Hnd, Text := Line);
  Line := CONCAT('end_ms=', UDINT_TO_STRING(RxMs1), TxCRLF); Ok := Ok AND TxLogPut(Hnd := Hnd, Text := Line);
  Line := CONCAT('duration_ms=', UDINT_TO_STRING(RxDur), TxCRLF); Ok := Ok AND TxLogPut(Hnd := Hnd, Text := Line);
  Line := CONCAT('plc_cycles=', UDINT_TO_STRING(RxCycN), TxCRLF); Ok := Ok AND TxLogPut(Hnd := Hnd, Text := Line);
  Line := CONCAT('committed=', BOOL_TO_STRING(RxCommitted), TxCRLF); Ok := Ok AND TxLogPut(Hnd := Hnd, Text := Line);
  IF RxWorkErr = 0 THEN Line := CONCAT('result=OK', TxCRLF);
  ELSE Line := CONCAT('result=ERROR', TxCRLF);
  END_IF;
  Ok := Ok AND TxLogPut(Hnd := Hnd, Text := Line);
  Line := CONCAT('error=', USINT_TO_STRING(RxWorkErr), TxCRLF); Ok := Ok AND TxLogPut(Hnd := Hnd, Text := Line);
  Line := CONCAT('error_text=', RxErrTxt, TxCRLF); Ok := Ok AND TxLogPut(Hnd := Hnd, Text := Line);
  Closed := FileClose(hFile := Hnd);
  RxWriteLog := Ok AND Closed;
END_FUNCTION

// Spracuje jednu položku parsera JSON: hlavičku, číslo vety alebo hodnotu poľa. ; Process one JSON parser item: header, record number, or field value.
// Porovná názvy JSON s presnou cestou schémy a odmieta neznáme alebo duplicitné polia. ; Match JSON names against schema paths and reject unknown or duplicate fields.
FUNCTION RxProcessItem : BOOL
  VAR
    Name     : STRING[255];  // Názov práve spracúvanej položky JSON ; Name of the JSON item currently being processed
    Value    : STRING[255];  // Hodnota načítaná z JSON parsera ; Value read from the JSON parser
    Expected : STRING[255];  // Očakávaný názov nasledujúceho poľa ; Expected name of the next field
    NextIdx  : UINT;         // Index nasledujúcej položky parsera ; Index of the next parser item
    Lf       : UINT;         // Index cieľového poľa v schéme ; Target leaf-field index in the schema
    LastLf   : UINT;         // Posledný index poľa v schéme typu ; Last leaf-field index for the type
    Pos      : UDINT;        // Adresa alebo pozícia hodnoty v pracovnej pamäti ; Address or position of the value in staging memory
    Found    : BOOL;         // Príznak nájdenia poľa v schéme ; Flag indicating that the field was found in the schema
  END_VAR
  RxProcessItem := FALSE;
  Name := RxInfo.item.name;
  Value := RxInfo.item.value;
  RxLastName := Name;

  IF Name = 'rq' THEN RxFileRq := STRING_TO_UDINT(Value); RxProcessItem := TRUE; RETURN; END_IF;
  IF Name = 'cf' THEN RxCfW := STRING_TO_USINT(Value); RxHdrCf := TRUE; RxProcessItem := TRUE; RETURN; END_IF;
  IF Name = 'type' THEN RxTypeW := Value; RxHdrType := TRUE; RxProcessItem := TRUE; RETURN; END_IF;
  IF Name = 'from' THEN RxFrom := STRING_TO_UDINT(Value); RxHdrFrom := TRUE; RxProcessItem := TRUE; RETURN; END_IF;
  IF Name = 'to' THEN RxTo := STRING_TO_UDINT(Value); RxHdrTo := TRUE; RxProcessItem := TRUE; RETURN; END_IF;
  IF Name = 'count' THEN RxCount := STRING_TO_UDINT(Value); RxHdrCount := TRUE; RxProcessItem := TRUE; RETURN; END_IF;

  NextIdx := RxIdx;
  IF RxHaveRec THEN NextIdx := RxIdx + 1; END_IF;
  Expected := CONCAT('data[', UINT_TO_STRING(NextIdx), '].rec');
  // Začiatok novej vety uzavrie predchádzajúcu a overí jej úplnosť. ; A new record marker closes the previous record and checks its completeness.
  IF Name = Expected THEN
    IF RxHaveRec THEN
      IF RxFieldsCur <> aSch[RxCfW].LCnt THEN RxWorkErr := 4; RxErrTxt := 'Missing fields in record'; RETURN; END_IF;
      RxRecordsDone := RxRecordsDone + 1;
      RxIdx := NextIdx;
    ELSE
      IF NOT RxPrepare() THEN RETURN; END_IF;
      RxIdx := 0;
    END_IF;
    IF RxIdx >= UDINT_TO_UINT(RxCount) THEN RxWorkErr := 4; RxErrTxt := 'Too many records'; RETURN; END_IF;
    RxRecCur := STRING_TO_UDINT(Value);
    IF RxRecCur <> RxFrom + UINT_TO_UDINT(RxIdx) THEN RxWorkErr := 4; RxErrTxt := 'Record number mismatch'; RETURN; END_IF;
    FOR Lf := 1 TO SCH_LEAF_N DO RxLeafSeen[Lf] := FALSE; END_FOR;
    RxFieldsCur := 0;
    RxHaveRec := TRUE;
    RxProcessItem := TRUE;
    RETURN;
  END_IF;

  IF NOT RxHaveRec OR NOT RxPrepared THEN RxWorkErr := 4; RxErrTxt := 'Data before record header'; RETURN; END_IF;
  LastLf := aSch[RxCfW].LFst + aSch[RxCfW].LCnt - 1;
  // Hľadá presnú cestu poľa v rozsahu listov vybranej schémy. ; Search for the exact field path within the selected schema's leaf range.
  FOR Lf := aSch[RxCfW].LFst TO LastLf DO
    Expected := CONCAT('data[', UINT_TO_STRING(RxIdx), '].value.', aLeaf[Lf].Pth);
    IF Name = Expected THEN
      Found := TRUE;
      IF RxLeafSeen[Lf] THEN RxWorkErr := 5; RxErrTxt := 'Duplicate field'; RETURN; END_IF;
      Pos := PTR_TO_UDINT(ADR(RxTmp[0])) + (RxRecCur - RxFrom) * aSch[RxCfW].Siz + UINT_TO_UDINT(aLeaf[Lf].Ofs);
      IF Pos + UINT_TO_UDINT(aLeaf[Lf].Span) > PTR_TO_UDINT(ADR(RxTmp[0])) + RxStageBytes THEN
        RxWorkErr := 6; RxErrTxt := 'Field outside staging'; RETURN;
      END_IF;
      IF NOT RxSetValue(Lf := Lf, Pos := Pos, Value := Value) THEN RETURN; END_IF;
      RxLeafSeen[Lf] := TRUE;
      RxFieldsCur := RxFieldsCur + 1;
      RxFieldsDone := RxFieldsDone + 1;
      RxProcessItem := TRUE;
      RETURN;
    END_IF;
  END_FOR;
  IF NOT Found THEN RxWorkErr := 5; RxErrTxt := 'Unknown JSON field'; END_IF;
END_FUNCTION

// Skontroluje úplnosť importu a až potom prenesie pripravené dáta do mRam. ; Verify import completeness and only then copy staged data into mRam.
// Commit do mRam nastane až po kontrole poslednej vety a všetkých povinných polí. ; Commit to mRam occurs only after checking the last record and all required fields.
FUNCTION RxEnd : BOOL
  VAR
    Copied : UDINT;  // Počet bajtov skopírovaných do pracovnej pamäte ; Number of bytes copied to staging memory
    LogOk  : BOOL;   // Výsledok zápisu meracieho logu ; Result of writing the measurement log
  END_VAR
  RxCommitted := FALSE;
  IF RxWorkErr = 0 THEN
    IF NOT RxPrepared OR NOT RxHaveRec OR (RxFieldsCur <> aSch[RxCfW].LCnt) THEN
      RxWorkErr := 4; RxErrTxt := 'Incomplete final record';
    ELSE
      RxRecordsDone := RxRecordsDone + 1;
      IF RxRecordsDone <> RxCount THEN RxWorkErr := 4; RxErrTxt := 'Record count mismatch'; END_IF;
    END_IF;
  END_IF;
  IF RxWorkErr = 0 THEN
    Copied := MemCpyPtr(source := ADR(RxTmp[0]),
      dest := UDINT_TO_PTR(aCfg[RxCfW].Ram + (RxFrom - 1) * aSch[RxCfW].Siz),
      length := RxStageBytes);
    IF Copied <> RxStageBytes THEN RxWorkErr := 7; RxErrTxt := 'mRam commit failed';
    ELSE RxCommitted := TRUE;
    END_IF;
  END_IF;
  RxMs1 := TxClockMs();
  RxDur := RxMs1 - RxMs0;
  RxCycN := RxCyc - RxCyc0 + 1;
  LogOk := RxWriteLog();
  IF (RxWorkErr = 0) AND NOT LogOk THEN RxWorkErr := 8; RxErrTxt := 'rx.log write failed'; END_IF;
  RxErr := RxWorkErr;
  RxDone := RxRqW;
  RxSt := 0;
  RxEnd := RxWorkErr = 0;
END_FUNCTION

// Vynuluje stav jednej požiadavky importu a spustí parser. ; Reset one import request's state and start the parser.
// Vynuluje počítadlá a príznaky, aby sa požiadavky navzájom nekontaminovali. ; Reset counters and flags so requests cannot contaminate one another.
FUNCTION RxStart : BOOL
  VAR
    Lf : UINT;  // Index cieľového poľa v schéme ; Target leaf-field index in the schema
  END_VAR
  RxRqW := RxRq;
  RxWorkErr := 0;
  RxErrTxt := '';
  RxLastName := '';
  RxCfW := 0;
  RxTypeW := '';
  RxFrom := 0;
  RxTo := 0;
  RxCount := 0;
  RxFileRq := 0;
  RxHdrCf := FALSE;
  RxHdrType := FALSE;
  RxHdrFrom := FALSE;
  RxHdrTo := FALSE;
  RxHdrCount := FALSE;
  RxPrepared := FALSE;
  RxHaveRec := FALSE;
  RxIdx := 0;
  RxRecCur := 0;
  RxFieldsCur := 0;
  RxFieldsDone := 0;
  RxRecordsDone := 0;
  RxStageBytes := 0;
  RxCommitted := FALSE;
  RxMs0 := TxClockMs();
  RxCyc0 := RxCyc;
  RxErr := 1;
  FOR Lf := 1 TO SCH_LEAF_N DO RxLeafSeen[Lf] := FALSE; END_FOR;
  RxSt := 1;
  RxStart := TRUE;
END_FUNCTION

// Stavový automat parsovania, validácie a potvrdenia rx.json. ; State machine for parsing, validating, and acknowledging rx.json.
// Každý cyklus posunie parser ; dokončená položka sa spracuje a EOF uzavrie požiadavku. ; Advance the parser each cycle ; process completed items and finish the request at EOF.
FUNCTION RxCycle : BOOL
  VAR
    Ok : BOOL;  // Príznak úspešného dokončenia kroku ; Flag indicating the step completed successfully
  END_VAR
  RxCyc := RxCyc + 1;
  RxCycle := TRUE;
  IF RxSt = 0 THEN
    RxParser(exec := FALSE, fileName := RxPath, JsonInfo := RxInfo);
    IF (RxRq = 0) OR (RxRq = RxRqSeen) THEN RETURN; END_IF;
    RxRqSeen := RxRq;
    // Po blokovom prenose povoľ import až po zložení a overení celého súboru. ; After block transfer, allow import only when the complete file is assembled and validated.
    IF (RbRq <> 0) AND NOT RbReady THEN
      RxErr := 9;
      RxDone := RxRq;
      RETURN;
    END_IF;
    RxCycle := RxStart();
    RETURN;
  END_IF;

  IF RxSt <> 1 THEN RxWorkErr := 1; RxErrTxt := 'Invalid RX state'; RxCycle := RxEnd(); RETURN; END_IF;
  RxParser(exec := TRUE, fileName := RxPath, JsonInfo := RxInfo);
  IF RxParser.done THEN
    IF NOT RxProcessItem() THEN RxCycle := RxEnd(); RETURN; END_IF;
  END_IF;
  IF RxParser.err THEN
    RxWorkErr := 2;
    RxErrTxt := RxParser.errTxt;
    RxCycle := RxEnd();
    RETURN;
  END_IF;
  IF RxParser.eof THEN
    Ok := RxEnd();
    RxCycle := Ok;
  END_IF;
END_FUNCTION
